FUNCTION_BLOCK "FB_SatelliteUnit"   // FB4, SCL
{ S7_Optimized_Access := 'TRUE' }
VERSION : 0.1
// Generated frame v0.12; change the declaration, then regenerate.
// stored: AutoNumber true, IsIECCheckEnabled false, IsRetainMemResEnabled false, MemoryReserve 100, SetENOAutomatically false, UDAEnableTagReadback false
   VAR_INPUT
      Execute { ExternalWritable := 'False'} : Bool;
      Abort { ExternalWritable := 'False'} : Bool;
      Command { ExternalWritable := 'False'} : DInt;
      ParCmd { ExternalWritable := 'False'} : "ST_DeclarationParCmd";
      ParentIndex { ExternalAccessible := 'False'; ExternalVisible := 'False'; ExternalWritable := 'False'} : DInt;
      Startup { ExternalAccessible := 'False'; ExternalVisible := 'False'; ExternalWritable := 'False'} : Bool;
   END_VAR
   VAR_OUTPUT
      Busy { ExternalWritable := 'False'} : Bool;
      Done { ExternalWritable := 'False'} : Bool;
      Error { ExternalWritable := 'False'} : Bool;
      Aborted { ExternalWritable := 'False'} : Bool;
      Held { ExternalWritable := 'False'} : Bool;
      ErrorID { ExternalWritable := 'False'} : DWord;
      Timing { ExternalWritable := 'False'} : "ST_ModuleTiming";
      OutCmd { ExternalWritable := 'False'} : "ST_DeclarationOutCmd";
      OutImm { ExternalWritable := 'False'} : "ST_UnitProbeImm";
   END_VAR
   VAR_IN_OUT
      Hal : "ST_SatelliteUnitHal";
   END_VAR
   VAR
      Status { ExternalWritable := 'False'; S7_SetPoint := 'True'} : "ST_ModuleStatus";
      Core { ExternalAccessible := 'False'; ExternalVisible := 'False'; ExternalWritable := 'False'; S7_SetPoint := 'True'} : "FRK_Core";
      ParCfg { ExternalWritable := 'False'; S7_SetPoint := 'True'} : "ST_DeclarationParCfg";
      LatchedParCmd { ExternalAccessible := 'False'; ExternalVisible := 'False'; ExternalWritable := 'False'; S7_SetPoint := 'True'} : "ST_DeclarationParCmd";
      StateFlags { ExternalWritable := 'False'; S7_SetPoint := 'True'} : Array[1..12] of "ST_StateFlag";
      StateFlagCount { ExternalWritable := 'False'} : Int;
      StateTouched { ExternalAccessible := 'False'; ExternalVisible := 'False'; ExternalWritable := 'False'} : Array[1..12] of Bool;
      Device { ExternalAccessible := 'False'; ExternalVisible := 'False'; ExternalWritable := 'False'; S7_SetPoint := 'True'} : "ST_UnitProbeDevice";
      StationCfg { ExternalWritable := 'False'; S7_SetPoint := 'True'} : "ST_UnitProbeStationCfg";
      ConfigStageParCfg { ExternalAccessible := 'False'; ExternalVisible := 'False'; ExternalWritable := 'False'; S7_SetPoint := 'True'} : "ST_DeclarationParCfg";
      ConfigDefaultParCfg { ExternalAccessible := 'False'; ExternalVisible := 'False'; ExternalWritable := 'False'; S7_SetPoint := 'True'} : "ST_DeclarationParCfg";
      ConfigStageStationCfg { ExternalAccessible := 'False'; ExternalVisible := 'False'; ExternalWritable := 'False'; S7_SetPoint := 'True'} : "ST_UnitProbeStationCfg";
      ConfigDefaultStationCfg { ExternalAccessible := 'False'; ExternalVisible := 'False'; ExternalWritable := 'False'; S7_SetPoint := 'True'} : "ST_UnitProbeStationCfg";
      ConfigStaged { ExternalAccessible := 'False'; ExternalVisible := 'False'; ExternalWritable := 'False'} : Bool;
      Unit { ExternalAccessible := 'False'; ExternalVisible := 'False'; ExternalWritable := 'False'; S7_SetPoint := 'True'} : "FRK_Unit";
      HmiRequest { S7_SetPoint := 'True'} : "ST_HmiRequest";
      ModePolicy { ExternalAccessible := 'False'; ExternalVisible := 'False'; ExternalWritable := 'False'; S7_SetPoint := 'True'} : Array[0..6] of "ST_ModePolicy";
      Access { ExternalWritable := 'False'; S7_SetPoint := 'True'} : "FRK_Access";
      HmiResponse { ExternalWritable := 'False'; S7_SetPoint := 'True'} : "ST_HmiResponse";
      ConfigRev { ExternalWritable := 'False'} : UDInt;
      ConfigCursor { ExternalAccessible := 'False'; ExternalVisible := 'False'; ExternalWritable := 'False'; S7_SetPoint := 'True'} : "FRK_ConfigCursor";
      Part { ExternalWritable := 'False'; S7_SetPoint := 'True'} : "ST_PartContext";
      Decision { ExternalWritable := 'False'; S7_SetPoint := 'True'} : "ST_DecisionRequest";
      DecisionAnswer { ExternalWritable := 'False'} : Int;
      History { ExternalWritable := 'False'; S7_SetPoint := 'True'} : Array[1..16] of "ST_Diagnostic";
      HistoryHead { ExternalWritable := 'False'} : Int;
      AlarmLog { ExternalWritable := 'False'; S7_SetPoint := 'True'} : "FRK_AlarmLog";
      ModeActivePublished { ExternalWritable := 'False'} : DInt;
      RunningPublished { ExternalWritable := 'False'} : Bool;
      StopPendingPublished { ExternalWritable := 'False'} : Bool;
      SupportedModesPublished { ExternalWritable := 'False'} : Array[0..6] of Bool;
      GoodCount { ExternalWritable := 'False'} : UDInt;
      NokCount { ExternalWritable := 'False'} : UDInt;
      ReworkCount { ExternalWritable := 'False'} : UDInt;
      NokReason { ExternalWritable := 'False'} : DInt;
      Cell { ExternalWritable := 'False'; S7_SetPoint := 'True'} : "FB_DeclarationCell";
      Inner { ExternalWritable := 'False'; S7_SetPoint := 'True'} : "FB_InnerUnit";
   END_VAR
   VAR_TEMP
      InstancePath : WString[254];
      RouteMatched : Bool;
      ManualMatched : Bool;
   END_VAR
   VAR CONSTANT
      EXEC_READY : DInt := 0;
      MODULE_TIER : DInt := 1;
   END_VAR
BEGIN

   // ---- GENERATED: setup
   IF #Startup OR NOT #Core.Named THEN
       #InstancePath := GetInstancePath(size := 0);
       "FRK_SetIdentity"(Core := #Core,
                         Status := #Status,
                         InstancePath := #InstancePath,
                         ModuleType := 1,
                         TypeId := 4,
                         Capabilities := DWORD#16#00000000,
                         ParentIndex := #ParentIndex,
                         TypeKey := 'Fraktal.Test.Satellite');
   END_IF;
   IF #Startup THEN "FRK_CfgRestore_SatelliteUnit"(Core := #Core,
                                                       Status := #Status,
                                                       ParCfg := #ParCfg,
                                                       StationCfg := #StationCfg,
                                                       ConfigStageParCfg := #ConfigStageParCfg,
                                                       ConfigDefaultParCfg := #ConfigDefaultParCfg,
                                                       ConfigStageStationCfg := #ConfigStageStationCfg,
                                                       ConfigDefaultStationCfg := #ConfigDefaultStationCfg);
   END_IF;
   "FRK_StateSweep"(Flags := #StateFlags,
                    Count := #StateFlagCount,
                    Touched := #StateTouched,
                    Startup := #Startup);
   IF #Startup OR #ConfigRev = 0 THEN
       #ConfigRev := "FRK_ConfigRevision"(Previous := #ConfigRev);
   END_IF;
   #SupportedModesPublished[0] := TRUE;
   #SupportedModesPublished[1] := TRUE;
   #SupportedModesPublished[2] := TRUE;
   #SupportedModesPublished[3] := FALSE;
   #SupportedModesPublished[4] := FALSE;
   #SupportedModesPublished[5] := FALSE;
   #SupportedModesPublished[6] := FALSE;
   "FRK_UnitPrepare"(Core := #Core,
                     Unit := #Unit,
                     Policy := #ModePolicy,
                     Request := #HmiRequest,
                     Response := #HmiResponse,
                     Startup := #Startup,
                     InitialMode := 1);
   "FRK_AlarmBegin"(AlarmLog := #AlarmLog,
                    Startup := #Startup);
   "FRK_AlarmHistoryBoot"(AlarmLog := #AlarmLog,
                          Startup := #Startup,
                          Scope := #Status.Name);
   "FRK_AccessPolicyBoot"(Access := #Access,
                          Startup := #Startup,
                          Root := #Core.ParentIndex = 0,
                          Scope := #Status.Name);
   "FRK_AccessCyclic"(Access := #Access,
                      Startup := #Startup,
                      SourcePath := STRING_TO_WSTRING(#Status.Name),
                      AlarmLog := #AlarmLog,
                      Revision := #ConfigRev);
   "FRK_UnitMailbox"(Core := #Core,
                     Unit := #Unit,
                     Status := #Status,
                     Policy := #ModePolicy,
                     Access := #Access,
                     Request := #HmiRequest,
                     Response := #HmiResponse,
                     Supported := #SupportedModesPublished);
   #Unit.ConfigBlocked := #Access.PolicyLost;
   // ---- GENERATED: begin
   "FRK_Begin"(Core := #Core,
               Status := #Status,
               Execute := #Unit.RunReq,
               Abort := (#Abort OR #Unit.AbortReq),
               Command := 1);
   IF #Core.EvCommandStart THEN
       #LatchedParCmd := #ParCmd;
       CASE #Core.Command OF
           1:
               "FRK_UnitRunStart"(Core := #Core,
                                  Status := #Status,
                                  Timeout := #ParCfg.Timeout,
                                  Label := 'Run');
           ELSE
               "FRK_Start"(Core := #Core,
                           Status := #Status,
                           Supported := FALSE,
                           Timeout := T#0ms,
                           Label := '');
       END_CASE;
   END_IF;
   IF #Core.EvCommandStart THEN
       // ---- AUTHORED: CommandStart
       #Device.Received := "FRK_PartReceived"(Core := #Core, Unit := #Unit, Status := #Status, Part := #Part, AlarmLog := #AlarmLog);
       IF #Device.Received THEN
           "FRK_PartStarted"(Unit := #Unit,
                             Status := #Status,
                             Part := #Part,
                             AlarmLog := #AlarmLog);
       END_IF;
       // ---- GENERATED: reaction end
   END_IF;
   // ---- AUTHORED: cyclic management
   IF #Hal.Cell.Clamp.BackgroundFault THEN
       "FRK_Fault"(Core := #Core,
                   Status := #Status,
                   ReasonCode := 2901,
                   Description := WSTRING#'test.unit.condition');
   END_IF;
   // ---- GENERATED: end management
   "FRK_Release_SatelliteUnit"(Unit := #Unit,
                               Hal := #Hal);
   IF #Core.RegIndex > 0 THEN
       "FRK_Registry".Rows[#Core.RegIndex].AlarmBlocking := #AlarmLog.Blocking;
   END_IF;
   #Unit.AlarmBlocking := "FRK_AlarmTreeBlocking"(Owner := #Core.RegIndex);
   "FRK_UnitConsume"(Core := #Core,
                     Unit := #Unit,
                     Status := #Status,
                     Policy := #ModePolicy,
                     Access := #Access,
                     Response := #HmiResponse,
                     Supported := #SupportedModesPublished);
   "FRK_UnitMode"(Core := #Core,
                  Unit := #Unit);
   IF #Core.EvModeExit THEN
       // ---- AUTHORED: ModeExit
       #Device.ExitCalls := #Device.ExitCalls + 1;
       IF #Hal.Cell.Clamp.ExitHold THEN
           #Core.HookResult := 1;
       ELSE
           #Core.HookResult := 0;
       END_IF;
       // ---- GENERATED: reaction end
   END_IF;
   "FRK_UnitModeResolve"(Core := #Core,
                         Unit := #Unit,
                         Status := #Status,
                         Policy := #ModePolicy,
                         Timeout := #ParCfg.Timeout);
   IF #Core.EvModeChanged THEN
       // ---- AUTHORED: ModeChanged
       #Device.Changes := #Device.Changes + 1;
       // ---- GENERATED: reaction end
   END_IF;
   "FRK_DecisionCyclic"(Owner := #Core.RegIndex,
                        Busy := #Core.Exec = 1,
                        Reset := #Startup OR #Unit.EvReset OR #Core.EvModeChanged,
                        AlarmLog := #AlarmLog);
   "FRK_UnitFollow"(Core := #Core,
                    Unit := #Unit,
                    Status := #Status,
                    Policy := #ModePolicy,
                    Access := #Access,
                    Supported := #SupportedModesPublished);
   IF #Unit.RequestPending AND (#Unit.Request.Kind = 11 OR #Unit.Request.Kind = 16) THEN
       #ManualMatched := FALSE;
       #RouteMatched := "FRK_Route_DeclarationCell"(Module := #Cell, Hal := #Hal.Cell, Request := #Unit.Request, Report := #HmiResponse.Report);
       #ManualMatched := #ManualMatched OR #RouteMatched;
       #RouteMatched := "FRK_Route_InnerUnit"(Module := #Inner, Hal := #Hal.Inner, Request := #Unit.Request, Report := #HmiResponse.Report);
       #ManualMatched := #ManualMatched OR #RouteMatched;
       IF NOT #ManualMatched THEN
           "FRK_ReleaseReason"(Report := #HmiResponse.Report,
                               Description := WSTRING#'std.error.unsupportedHmiRequest',
                               Reason := 2008,
                               Path := #Unit.Request.TargetPath,
                               Kind := 4);
       END_IF;
       #HmiResponse.Accepted := #Unit.Request.Kind = 16 OR #HmiResponse.Report.Released;
       IF #Unit.Request.Kind = 11 THEN
           IF #HmiResponse.Accepted THEN
               #HmiResponse.Diagnostic := WSTRING#'std.audit.manualCommandAccepted';
           ELSE
               #HmiResponse.Diagnostic := WSTRING#'std.audit.manualCommandRejected';
           END_IF;
       END_IF;
   END_IF;
   IF #Unit.EvReset THEN
       "FRK_AlarmOperatorReset"(AlarmLog := #AlarmLog);
   END_IF;
   IF #Unit.EvReset THEN
       // ---- AUTHORED: OperatorReset
       #Device.Resets := #Device.Resets + 1;
       // ---- GENERATED: reset reaction end
   END_IF;
   IF #Core.ReleasePending OR #Unit.ReleaseChildren THEN
       "FRK_ReleaseCommand"(Core := #Cell.Core,
                            Execute := #Cell.Execute);
       "FRK_ReleaseCommand"(Core := #Inner.Core,
                            Execute := #Inner.Execute);
   END_IF;
   // ---- GENERATED: child call
   #Cell(ParentIndex := #Core.RegIndex,
         Startup := #Startup,
         Hal := #Hal.Cell);
   "FRK_ManualFinish"(Core := #Cell.Core,
                      Execute := #Cell.Execute,
                      ManualOwned := #Cell.ManualOwned);
   "FRK_UnitCascade"(ParentUnit := #Unit,
                     Core := #Inner.Core,
                     Unit := #Inner.Unit,
                     Status := #Inner.Status,
                     Policy := #Inner.ModePolicy,
                     Access := #Inner.Access,
                     Supported := #Inner.SupportedModesPublished,
                     AlarmLog := #AlarmLog);
   // ---- GENERATED: child call
   #Inner(ParentIndex := #Core.RegIndex,
          Startup := #Startup,
          Hal := #Hal.Inner);
   #Unit.CascadePending := FALSE;
   IF #Unit.RequestPending AND #Unit.Request.Kind = 23 THEN
       #HmiResponse.Accepted := FALSE;
       #HmiResponse.Report.Count := 0;
       #HmiResponse.Report.Released := TRUE;
       #HmiResponse.Diagnostic := WSTRING#'';
       "FRK_ConfigBegin"(Cursor := #ConfigCursor,
                         Page := #HmiResponse.ConfigPage,
                         PageIndex := #Unit.Request.IntValue,
                         Revision := #ConfigRev);
       IF #Unit.Request.DurationMs <> 0 THEN
           #HmiResponse.Diagnostic := WSTRING#'std.error.modelNotAvailable';
       ELSIF #Unit.Request.IntValue < 0 OR #Unit.Request.IntValue > 32767 THEN
           #HmiResponse.Diagnostic := WSTRING#'std.error.hmiRequestRejected';
       ELSE
           "FRK_ConfigUnit"(Scope := #Status.Name,
                            Policy := #ModePolicy,
                            ModelCount := 0,
                            ReadLevel := #Access.Policy.Required[0],
                            Readable := #Access.CurrentLevel >= #Access.Policy.Required[0],
                            Cursor := #ConfigCursor,
                            Page := #HmiResponse.ConfigPage);
           "FRK_Config_DeclarationCell"(Module := #Cell,
                                        Access := #Access,
                                        RootIndex := "FRK_ConfigRoot"(RegIndex := #Core.RegIndex),
                                        ModelIndex := 0,
                                        Cursor := #ConfigCursor,
                                        Page := #HmiResponse.ConfigPage);
           "FRK_Config_InnerUnit"(Module := #Inner,
                                  Access := #Access,
                                  RootIndex := "FRK_ConfigRoot"(RegIndex := #Core.RegIndex),
                                  ModelIndex := 0,
                                  Cursor := #ConfigCursor,
                                  Page := #HmiResponse.ConfigPage);
           "FRK_ConfigFinish"(Cursor := #ConfigCursor,
                              Page := #HmiResponse.ConfigPage);
           #HmiResponse.Accepted := TRUE;
       END_IF;
   END_IF;
   "FRK_RouteAbort"(Core := #Core,
                    Abort := (#Abort OR #Unit.AbortReq));
   IF #Core.EvAbort THEN
       "FRK_PartAborted"(Core := #Core,
                         Unit := #Unit,
                         Status := #Status,
                         Part := #Part,
                         AlarmLog := #AlarmLog);
   END_IF;
   IF #Core.Dispatch AND #Core.RegIndex > 0 AND NOT "FRK_Registry".Fault THEN
       // ---- AUTHORED: dispatch
       IF #Hal.Cell.Clamp.Finish THEN
           #Device.Processed := FALSE;
           IF #Unit.CarrierIndex = 0 THEN
               #Device.Processed := TRUE;
           ELSE
               #Device.Processed := "FRK_PartProcessed"(Core := #Core, Unit := #Unit, Status := #Status, Part := #Part, AlarmLog := #AlarmLog, Verdict := #Hal.Cell.Clamp.Verdict, Reason := #Hal.Cell.Clamp.Diag.ReasonCode);
           END_IF;
           IF #Device.Processed THEN
               #Device.Cycles := #Device.Cycles + 1;
               IF #Unit.StopReq THEN
                   "FRK_Complete"(Core := #Core,
                                  Status := #Status);
               ELSE
                   #Device.Received := "FRK_PartReceived"(Core := #Core, Unit := #Unit, Status := #Status, Part := #Part, AlarmLog := #AlarmLog);
                   IF #Device.Received THEN
                       "FRK_PartStarted"(Unit := #Unit,
                                         Status := #Status,
                                         Part := #Part,
                                         AlarmLog := #AlarmLog);
                   END_IF;
               END_IF;
           END_IF;
       END_IF;
       // ---- GENERATED: end dispatch
   END_IF;
   "FRK_End"(Core := #Core,
             Status := #Status,
             Busy => #Busy,
             Done => #Done,
             Error => #Error,
             Aborted => #Aborted,
             Held => #Held,
             ErrorID => #ErrorID,
             Timing => #Timing);
   "FRK_DecisionCyclic"(Owner := #Core.RegIndex,
                        Busy := #Core.Exec = 1,
                        Reset := #Startup OR #Unit.EvReset OR #Core.EvModeChanged,
                        AlarmLog := #AlarmLog);
   "FRK_DecisionPublish"(Owner := #Core.RegIndex,
                         Decision := #Decision,
                         DecisionAnswer := #DecisionAnswer);
   IF NOT #Unit.EvReset THEN
       "FRK_AlarmCapture"(AlarmLog := #AlarmLog,
                          Core := #Core,
                          Status := #Status);
       "FRK_Capture_DeclarationCell"(Module := #Cell,
                                     AlarmLog := #AlarmLog);
       "FRK_AlarmEnd"(AlarmLog := #AlarmLog);
   END_IF;
   IF #Core.RegIndex > 0 THEN
       "FRK_Registry".Rows[#Core.RegIndex].AlarmBlocking := #AlarmLog.Blocking;
   END_IF;
   #Unit.AlarmBlocking := "FRK_AlarmTreeBlocking"(Owner := #Core.RegIndex);
   "FRK_AccessPersist"(Access := #Access,
                       Unit := #Unit,
                       Response := #HmiResponse,
                       SourcePath := STRING_TO_WSTRING(#Status.Name),
                       AlarmLog := #AlarmLog);
   "FRK_AccessFinish"(Access := #Access,
                      Unit := #Unit,
                      Response := #HmiResponse,
                      SourcePath := STRING_TO_WSTRING(#Status.Name),
                      AlarmLog := #AlarmLog,
                      Revision := #ConfigRev);
   "FRK_UnitFinish"(Core := #Core,
                    Unit := #Unit,
                    Response := #HmiResponse,
                    Status := #Status,
                    Part := #Part,
                    AlarmLog := #AlarmLog,
                    History := #History,
                    Head := #HistoryHead);
   #ModeActivePublished := #Unit.Mode;
   #RunningPublished := #Core.Exec = 1;
   #StopPendingPublished := #Unit.StopReq AND #Core.Exec = 1;
   #GoodCount := #Unit.Good;
   #NokCount := #Unit.Nok;
   #ReworkCount := #Unit.Rework;
   #NokReason := #Unit.NokReason;
   // ---- AUTHORED: unconditional cyclic/derived data
   #OutImm.Cycles := #Device.Cycles;
   #OutImm.ExitCalls := #Device.ExitCalls;
   #OutImm.Changes := #Device.Changes;
   #OutImm.Resets := #Device.Resets;
   #OutImm.AtHome := "FRK_State"(Idx := 1, Key := 'project.state.atHome', Ok := #Hal.Cell.Clamp.Sample = 0, Flags := #StateFlags, Count := #StateFlagCount, Touched := #StateTouched);
   // ---- GENERATED: frame end
END_FUNCTION_BLOCK

FUNCTION_BLOCK "FB_InnerUnit"   // FB3, SCL
{ S7_Optimized_Access := 'TRUE' }
VERSION : 0.1
// Generated frame v0.12; change the declaration, then regenerate.
// stored: AutoNumber true, IsIECCheckEnabled false, IsRetainMemResEnabled false, MemoryReserve 100, SetENOAutomatically false, UDAEnableTagReadback false
   VAR_INPUT
      Execute { ExternalWritable := 'False'} : Bool;
      Abort { ExternalWritable := 'False'} : Bool;
      Command { ExternalWritable := 'False'} : DInt;
      ParCmd { ExternalWritable := 'False'} : "ST_DeclarationParCmd";
      ParentIndex { ExternalAccessible := 'False'; ExternalVisible := 'False'; ExternalWritable := 'False'} : DInt;
      Startup { ExternalAccessible := 'False'; ExternalVisible := 'False'; ExternalWritable := 'False'} : Bool;
   END_VAR
   VAR_OUTPUT
      Busy { ExternalWritable := 'False'} : Bool;
      Done { ExternalWritable := 'False'} : Bool;
      Error { ExternalWritable := 'False'} : Bool;
      Aborted { ExternalWritable := 'False'} : Bool;
      Held { ExternalWritable := 'False'} : Bool;
      ErrorID { ExternalWritable := 'False'} : DWord;
      Timing { ExternalWritable := 'False'} : "ST_ModuleTiming";
      OutCmd { ExternalWritable := 'False'} : "ST_DeclarationOutCmd";
      OutImm { ExternalWritable := 'False'} : "ST_UnitProbeImm";
   END_VAR
   VAR_IN_OUT
      Hal : "ST_InnerUnitHal";
   END_VAR
   VAR
      Status { ExternalWritable := 'False'; S7_SetPoint := 'True'} : "ST_ModuleStatus";
      Core { ExternalAccessible := 'False'; ExternalVisible := 'False'; ExternalWritable := 'False'; S7_SetPoint := 'True'} : "FRK_Core";
      ParCfg { ExternalWritable := 'False'; S7_SetPoint := 'True'} : "ST_DeclarationParCfg";
      LatchedParCmd { ExternalAccessible := 'False'; ExternalVisible := 'False'; ExternalWritable := 'False'; S7_SetPoint := 'True'} : "ST_DeclarationParCmd";
      StateFlags { ExternalWritable := 'False'; S7_SetPoint := 'True'} : Array[1..12] of "ST_StateFlag";
      StateFlagCount { ExternalWritable := 'False'} : Int;
      StateTouched { ExternalAccessible := 'False'; ExternalVisible := 'False'; ExternalWritable := 'False'} : Array[1..12] of Bool;
      Device { ExternalAccessible := 'False'; ExternalVisible := 'False'; ExternalWritable := 'False'; S7_SetPoint := 'True'} : "ST_UnitProbeDevice";
      StationCfg { ExternalWritable := 'False'; S7_SetPoint := 'True'} : "ST_UnitProbeStationCfg";
      ConfigStageParCfg { ExternalAccessible := 'False'; ExternalVisible := 'False'; ExternalWritable := 'False'; S7_SetPoint := 'True'} : "ST_DeclarationParCfg";
      ConfigDefaultParCfg { ExternalAccessible := 'False'; ExternalVisible := 'False'; ExternalWritable := 'False'; S7_SetPoint := 'True'} : "ST_DeclarationParCfg";
      ConfigStageStationCfg { ExternalAccessible := 'False'; ExternalVisible := 'False'; ExternalWritable := 'False'; S7_SetPoint := 'True'} : "ST_UnitProbeStationCfg";
      ConfigDefaultStationCfg { ExternalAccessible := 'False'; ExternalVisible := 'False'; ExternalWritable := 'False'; S7_SetPoint := 'True'} : "ST_UnitProbeStationCfg";
      ConfigStaged { ExternalAccessible := 'False'; ExternalVisible := 'False'; ExternalWritable := 'False'} : Bool;
      Unit { ExternalAccessible := 'False'; ExternalVisible := 'False'; ExternalWritable := 'False'; S7_SetPoint := 'True'} : "FRK_Unit";
      HmiRequest { S7_SetPoint := 'True'} : "ST_HmiRequest";
      ModePolicy { ExternalAccessible := 'False'; ExternalVisible := 'False'; ExternalWritable := 'False'; S7_SetPoint := 'True'} : Array[0..6] of "ST_ModePolicy";
      Access { ExternalWritable := 'False'; S7_SetPoint := 'True'} : "FRK_Access";
      HmiResponse { ExternalWritable := 'False'; S7_SetPoint := 'True'} : "ST_HmiResponse";
      ConfigRev { ExternalWritable := 'False'} : UDInt;
      ConfigCursor { ExternalAccessible := 'False'; ExternalVisible := 'False'; ExternalWritable := 'False'; S7_SetPoint := 'True'} : "FRK_ConfigCursor";
      Part { ExternalWritable := 'False'; S7_SetPoint := 'True'} : "ST_PartContext";
      Decision { ExternalWritable := 'False'; S7_SetPoint := 'True'} : "ST_DecisionRequest";
      DecisionAnswer { ExternalWritable := 'False'} : Int;
      History { ExternalWritable := 'False'; S7_SetPoint := 'True'} : Array[1..16] of "ST_Diagnostic";
      HistoryHead { ExternalWritable := 'False'} : Int;
      AlarmLog { ExternalWritable := 'False'; S7_SetPoint := 'True'} : "FRK_AlarmLog";
      ModeActivePublished { ExternalWritable := 'False'} : DInt;
      RunningPublished { ExternalWritable := 'False'} : Bool;
      StopPendingPublished { ExternalWritable := 'False'} : Bool;
      SupportedModesPublished { ExternalWritable := 'False'} : Array[0..6] of Bool;
      GoodCount { ExternalWritable := 'False'} : UDInt;
      NokCount { ExternalWritable := 'False'} : UDInt;
      ReworkCount { ExternalWritable := 'False'} : UDInt;
      NokReason { ExternalWritable := 'False'} : DInt;
      Cell { ExternalWritable := 'False'; S7_SetPoint := 'True'} : "FB_DeclarationCell";
   END_VAR
   VAR_TEMP
      InstancePath : WString[254];
      RouteMatched : Bool;
      ManualMatched : Bool;
   END_VAR
   VAR CONSTANT
      EXEC_READY : DInt := 0;
      MODULE_TIER : DInt := 1;
   END_VAR
BEGIN

   // ---- GENERATED: setup
   IF #Startup OR NOT #Core.Named THEN
       #InstancePath := GetInstancePath(size := 0);
       "FRK_SetIdentity"(Core := #Core,
                         Status := #Status,
                         InstancePath := #InstancePath,
                         ModuleType := 1,
                         TypeId := 5,
                         Capabilities := DWORD#16#00000000,
                         ParentIndex := #ParentIndex,
                         TypeKey := 'Fraktal.Test.Inner');
   END_IF;
   IF #Startup THEN "FRK_CfgRestore_InnerUnit"(Core := #Core,
                                                   Status := #Status,
                                                   ParCfg := #ParCfg,
                                                   StationCfg := #StationCfg,
                                                   ConfigStageParCfg := #ConfigStageParCfg,
                                                   ConfigDefaultParCfg := #ConfigDefaultParCfg,
                                                   ConfigStageStationCfg := #ConfigStageStationCfg,
                                                   ConfigDefaultStationCfg := #ConfigDefaultStationCfg);
   END_IF;
   "FRK_StateSweep"(Flags := #StateFlags,
                    Count := #StateFlagCount,
                    Touched := #StateTouched,
                    Startup := #Startup);
   IF #Startup OR #ConfigRev = 0 THEN
       #ConfigRev := "FRK_ConfigRevision"(Previous := #ConfigRev);
   END_IF;
   #SupportedModesPublished[0] := TRUE;
   #SupportedModesPublished[1] := TRUE;
   #SupportedModesPublished[2] := TRUE;
   #SupportedModesPublished[3] := FALSE;
   #SupportedModesPublished[4] := FALSE;
   #SupportedModesPublished[5] := FALSE;
   #SupportedModesPublished[6] := FALSE;
   "FRK_UnitPrepare"(Core := #Core,
                     Unit := #Unit,
                     Policy := #ModePolicy,
                     Request := #HmiRequest,
                     Response := #HmiResponse,
                     Startup := #Startup,
                     InitialMode := 1);
   "FRK_AlarmBegin"(AlarmLog := #AlarmLog,
                    Startup := #Startup);
   "FRK_AlarmHistoryBoot"(AlarmLog := #AlarmLog,
                          Startup := #Startup,
                          Scope := #Status.Name);
   "FRK_AccessPolicyBoot"(Access := #Access,
                          Startup := #Startup,
                          Root := #Core.ParentIndex = 0,
                          Scope := #Status.Name);
   "FRK_AccessCyclic"(Access := #Access,
                      Startup := #Startup,
                      SourcePath := STRING_TO_WSTRING(#Status.Name),
                      AlarmLog := #AlarmLog,
                      Revision := #ConfigRev);
   "FRK_UnitMailbox"(Core := #Core,
                     Unit := #Unit,
                     Status := #Status,
                     Policy := #ModePolicy,
                     Access := #Access,
                     Request := #HmiRequest,
                     Response := #HmiResponse,
                     Supported := #SupportedModesPublished);
   #Unit.ConfigBlocked := #Access.PolicyLost;
   // ---- GENERATED: begin
   "FRK_Begin"(Core := #Core,
               Status := #Status,
               Execute := #Unit.RunReq,
               Abort := (#Abort OR #Unit.AbortReq),
               Command := 1);
   IF #Core.EvCommandStart THEN
       #LatchedParCmd := #ParCmd;
       CASE #Core.Command OF
           1:
               "FRK_UnitRunStart"(Core := #Core,
                                  Status := #Status,
                                  Timeout := #ParCfg.Timeout,
                                  Label := 'Run');
           ELSE
               "FRK_Start"(Core := #Core,
                           Status := #Status,
                           Supported := FALSE,
                           Timeout := T#0ms,
                           Label := '');
       END_CASE;
   END_IF;
   IF #Core.EvCommandStart THEN
       // ---- AUTHORED: CommandStart
       #Device.Received := "FRK_PartReceived"(Core := #Core, Unit := #Unit, Status := #Status, Part := #Part, AlarmLog := #AlarmLog);
       IF #Device.Received THEN
           "FRK_PartStarted"(Unit := #Unit,
                             Status := #Status,
                             Part := #Part,
                             AlarmLog := #AlarmLog);
       END_IF;
       // ---- GENERATED: reaction end
   END_IF;
   // ---- AUTHORED: cyclic management
   IF #Hal.Cell.Clamp.BackgroundFault THEN
       "FRK_Fault"(Core := #Core,
                   Status := #Status,
                   ReasonCode := 2901,
                   Description := WSTRING#'test.unit.condition');
   END_IF;
   // ---- GENERATED: end management
   "FRK_Release_InnerUnit"(Unit := #Unit,
                           Hal := #Hal);
   IF #Core.RegIndex > 0 THEN
       "FRK_Registry".Rows[#Core.RegIndex].AlarmBlocking := #AlarmLog.Blocking;
   END_IF;
   #Unit.AlarmBlocking := "FRK_AlarmTreeBlocking"(Owner := #Core.RegIndex);
   "FRK_UnitConsume"(Core := #Core,
                     Unit := #Unit,
                     Status := #Status,
                     Policy := #ModePolicy,
                     Access := #Access,
                     Response := #HmiResponse,
                     Supported := #SupportedModesPublished);
   "FRK_UnitMode"(Core := #Core,
                  Unit := #Unit);
   IF #Core.EvModeExit THEN
       // ---- AUTHORED: ModeExit
       #Device.ExitCalls := #Device.ExitCalls + 1;
       IF #Hal.Cell.Clamp.ExitHold THEN
           #Core.HookResult := 1;
       ELSE
           #Core.HookResult := 0;
       END_IF;
       // ---- GENERATED: reaction end
   END_IF;
   "FRK_UnitModeResolve"(Core := #Core,
                         Unit := #Unit,
                         Status := #Status,
                         Policy := #ModePolicy,
                         Timeout := #ParCfg.Timeout);
   IF #Core.EvModeChanged THEN
       // ---- AUTHORED: ModeChanged
       #Device.Changes := #Device.Changes + 1;
       // ---- GENERATED: reaction end
   END_IF;
   "FRK_DecisionCyclic"(Owner := #Core.RegIndex,
                        Busy := #Core.Exec = 1,
                        Reset := #Startup OR #Unit.EvReset OR #Core.EvModeChanged,
                        AlarmLog := #AlarmLog);
   "FRK_UnitFollow"(Core := #Core,
                    Unit := #Unit,
                    Status := #Status,
                    Policy := #ModePolicy,
                    Access := #Access,
                    Supported := #SupportedModesPublished);
   IF #Unit.RequestPending AND (#Unit.Request.Kind = 11 OR #Unit.Request.Kind = 16) THEN
       #ManualMatched := FALSE;
       #RouteMatched := "FRK_Route_DeclarationCell"(Module := #Cell, Hal := #Hal.Cell, Request := #Unit.Request, Report := #HmiResponse.Report);
       #ManualMatched := #ManualMatched OR #RouteMatched;
       IF NOT #ManualMatched THEN
           "FRK_ReleaseReason"(Report := #HmiResponse.Report,
                               Description := WSTRING#'std.error.unsupportedHmiRequest',
                               Reason := 2008,
                               Path := #Unit.Request.TargetPath,
                               Kind := 4);
       END_IF;
       #HmiResponse.Accepted := #Unit.Request.Kind = 16 OR #HmiResponse.Report.Released;
       IF #Unit.Request.Kind = 11 THEN
           IF #HmiResponse.Accepted THEN
               #HmiResponse.Diagnostic := WSTRING#'std.audit.manualCommandAccepted';
           ELSE
               #HmiResponse.Diagnostic := WSTRING#'std.audit.manualCommandRejected';
           END_IF;
       END_IF;
   END_IF;
   IF #Unit.EvReset THEN
       "FRK_AlarmOperatorReset"(AlarmLog := #AlarmLog);
   END_IF;
   IF #Unit.EvReset THEN
       // ---- AUTHORED: OperatorReset
       #Device.Resets := #Device.Resets + 1;
       // ---- GENERATED: reset reaction end
   END_IF;
   IF #Core.ReleasePending OR #Unit.ReleaseChildren THEN
       "FRK_ReleaseCommand"(Core := #Cell.Core,
                            Execute := #Cell.Execute);
   END_IF;
   // ---- GENERATED: child call
   #Cell(ParentIndex := #Core.RegIndex,
         Startup := #Startup,
         Hal := #Hal.Cell);
   "FRK_ManualFinish"(Core := #Cell.Core,
                      Execute := #Cell.Execute,
                      ManualOwned := #Cell.ManualOwned);
   #Unit.CascadePending := FALSE;
   IF #Unit.RequestPending AND #Unit.Request.Kind = 23 THEN
       #HmiResponse.Accepted := FALSE;
       #HmiResponse.Report.Count := 0;
       #HmiResponse.Report.Released := TRUE;
       #HmiResponse.Diagnostic := WSTRING#'';
       "FRK_ConfigBegin"(Cursor := #ConfigCursor,
                         Page := #HmiResponse.ConfigPage,
                         PageIndex := #Unit.Request.IntValue,
                         Revision := #ConfigRev);
       IF #Unit.Request.DurationMs <> 0 THEN
           #HmiResponse.Diagnostic := WSTRING#'std.error.modelNotAvailable';
       ELSIF #Unit.Request.IntValue < 0 OR #Unit.Request.IntValue > 32767 THEN
           #HmiResponse.Diagnostic := WSTRING#'std.error.hmiRequestRejected';
       ELSE
           "FRK_ConfigUnit"(Scope := #Status.Name,
                            Policy := #ModePolicy,
                            ModelCount := 0,
                            ReadLevel := #Access.Policy.Required[0],
                            Readable := #Access.CurrentLevel >= #Access.Policy.Required[0],
                            Cursor := #ConfigCursor,
                            Page := #HmiResponse.ConfigPage);
           "FRK_Config_DeclarationCell"(Module := #Cell,
                                        Access := #Access,
                                        RootIndex := "FRK_ConfigRoot"(RegIndex := #Core.RegIndex),
                                        ModelIndex := 0,
                                        Cursor := #ConfigCursor,
                                        Page := #HmiResponse.ConfigPage);
           "FRK_ConfigFinish"(Cursor := #ConfigCursor,
                              Page := #HmiResponse.ConfigPage);
           #HmiResponse.Accepted := TRUE;
       END_IF;
   END_IF;
   "FRK_RouteAbort"(Core := #Core,
                    Abort := (#Abort OR #Unit.AbortReq));
   IF #Core.EvAbort THEN
       "FRK_PartAborted"(Core := #Core,
                         Unit := #Unit,
                         Status := #Status,
                         Part := #Part,
                         AlarmLog := #AlarmLog);
   END_IF;
   IF #Core.Dispatch AND #Core.RegIndex > 0 AND NOT "FRK_Registry".Fault THEN
       // ---- AUTHORED: dispatch
       IF #Hal.Cell.Clamp.Finish THEN
           #Device.Processed := FALSE;
           IF #Unit.CarrierIndex = 0 THEN
               #Device.Processed := TRUE;
           ELSE
               #Device.Processed := "FRK_PartProcessed"(Core := #Core, Unit := #Unit, Status := #Status, Part := #Part, AlarmLog := #AlarmLog, Verdict := #Hal.Cell.Clamp.Verdict, Reason := #Hal.Cell.Clamp.Diag.ReasonCode);
           END_IF;
           IF #Device.Processed THEN
               #Device.Cycles := #Device.Cycles + 1;
               IF #Unit.StopReq THEN
                   "FRK_Complete"(Core := #Core,
                                  Status := #Status);
               ELSE
                   #Device.Received := "FRK_PartReceived"(Core := #Core, Unit := #Unit, Status := #Status, Part := #Part, AlarmLog := #AlarmLog);
                   IF #Device.Received THEN
                       "FRK_PartStarted"(Unit := #Unit,
                                         Status := #Status,
                                         Part := #Part,
                                         AlarmLog := #AlarmLog);
                   END_IF;
               END_IF;
           END_IF;
       END_IF;
       // ---- GENERATED: end dispatch
   END_IF;
   "FRK_End"(Core := #Core,
             Status := #Status,
             Busy => #Busy,
             Done => #Done,
             Error => #Error,
             Aborted => #Aborted,
             Held => #Held,
             ErrorID => #ErrorID,
             Timing => #Timing);
   "FRK_DecisionCyclic"(Owner := #Core.RegIndex,
                        Busy := #Core.Exec = 1,
                        Reset := #Startup OR #Unit.EvReset OR #Core.EvModeChanged,
                        AlarmLog := #AlarmLog);
   "FRK_DecisionPublish"(Owner := #Core.RegIndex,
                         Decision := #Decision,
                         DecisionAnswer := #DecisionAnswer);
   IF NOT #Unit.EvReset THEN
       "FRK_AlarmCapture"(AlarmLog := #AlarmLog,
                          Core := #Core,
                          Status := #Status);
       "FRK_Capture_DeclarationCell"(Module := #Cell,
                                     AlarmLog := #AlarmLog);
       "FRK_AlarmEnd"(AlarmLog := #AlarmLog);
   END_IF;
   IF #Core.RegIndex > 0 THEN
       "FRK_Registry".Rows[#Core.RegIndex].AlarmBlocking := #AlarmLog.Blocking;
   END_IF;
   #Unit.AlarmBlocking := "FRK_AlarmTreeBlocking"(Owner := #Core.RegIndex);
   "FRK_AccessPersist"(Access := #Access,
                       Unit := #Unit,
                       Response := #HmiResponse,
                       SourcePath := STRING_TO_WSTRING(#Status.Name),
                       AlarmLog := #AlarmLog);
   "FRK_AccessFinish"(Access := #Access,
                      Unit := #Unit,
                      Response := #HmiResponse,
                      SourcePath := STRING_TO_WSTRING(#Status.Name),
                      AlarmLog := #AlarmLog,
                      Revision := #ConfigRev);
   "FRK_UnitFinish"(Core := #Core,
                    Unit := #Unit,
                    Response := #HmiResponse,
                    Status := #Status,
                    Part := #Part,
                    AlarmLog := #AlarmLog,
                    History := #History,
                    Head := #HistoryHead);
   #ModeActivePublished := #Unit.Mode;
   #RunningPublished := #Core.Exec = 1;
   #StopPendingPublished := #Unit.StopReq AND #Core.Exec = 1;
   #GoodCount := #Unit.Good;
   #NokCount := #Unit.Nok;
   #ReworkCount := #Unit.Rework;
   #NokReason := #Unit.NokReason;
   // ---- AUTHORED: unconditional cyclic/derived data
   #OutImm.Cycles := #Device.Cycles;
   #OutImm.ExitCalls := #Device.ExitCalls;
   #OutImm.Changes := #Device.Changes;
   #OutImm.Resets := #Device.Resets;
   #OutImm.AtHome := "FRK_State"(Idx := 1, Key := 'project.state.atHome', Ok := #Hal.Cell.Clamp.Sample = 0, Flags := #StateFlags, Count := #StateFlagCount, Touched := #StateTouched);
   // ---- GENERATED: frame end
END_FUNCTION_BLOCK

FUNCTION "FRK_AccessAudit" : Void   // FC53, SCL
{ S7_Optimized_Access := 'TRUE' }
VERSION : 0.1
// stored: AutoNumber true, IsIECCheckEnabled false, SetENOAutomatically false, UDAEnableTagReadback false
   VAR_INPUT
      What : WString;
      Who : String;
      SourcePath : WString;
   END_VAR
   VAR_IN_OUT
      AlarmLog : "FRK_AlarmLog";
   END_VAR
   VAR_TEMP
      Description : WString[480];
   END_VAR
BEGIN

   #Description := CONCAT(IN1 := #What, IN2 := WSTRING#': ');
   #Description := CONCAT(IN1 := #Description, IN2 := STRING_TO_WSTRING(#Who));
   "FRK_AlarmMessage"(AlarmLog := #AlarmLog,
                      Reason := 0,
                      Description := #Description,
                      SourcePath := #SourcePath);
END_FUNCTION

FUNCTION "FRK_AccessCancel" : Void   // FC48, SCL
{ S7_Optimized_Access := 'TRUE' }
VERSION : 0.1
// stored: AutoNumber true, IsIECCheckEnabled false, SetENOAutomatically false, UDAEnableTagReadback false
   VAR_IN_OUT
      Access : "FRK_Access";
   END_VAR
   VAR_TEMP
      Index : DInt;
   END_VAR
BEGIN

   #Access.LoginBusy := FALSE;
   #Access.CandidateUser := '';
   #Access.CandidateLevel := 0;
   #Access.Round := 0;
   FOR #Index := 0 TO 15 DO
       #Access.Salt[#Index] := 0;
   END_FOR;
   FOR #Index := 0 TO 31 DO
       #Access.Digest[#Index] := 0;
       #Access.Expected[#Index] := 0;
   END_FOR;
END_FUNCTION

FUNCTION "FRK_AccessCyclic" : Void   // FC54, SCL
{ S7_Optimized_Access := 'TRUE' }
VERSION : 0.1
// stored: AutoNumber true, IsIECCheckEnabled false, SetENOAutomatically false, UDAEnableTagReadback false
   VAR_INPUT
      Startup : Bool;
      SourcePath : WString;
   END_VAR
   VAR_IN_OUT
      Access : "FRK_Access";
      AlarmLog : "FRK_AlarmLog";
      Revision : UDInt;
   END_VAR
   VAR_TEMP
      Data : Array[0..47] of Byte;
      Index : DInt;
      Difference : Byte;
      HashOk : Bool;
   END_VAR
BEGIN

   #Access.LoginTimeoutMs := 6000;
   IF #Startup THEN
       "FRK_AccessLogout"(Access := #Access);
       #Access.LoginResultSequence := 0;
   END_IF;
   IF #Access.ProviderGeneration <> "FRK_LocalUsers".Generation OR NOT "FRK_AccessStorage".UsersReady THEN
       IF #Access.CurrentLevel > 0 THEN
           "FRK_AccessAudit"(AlarmLog := #AlarmLog,
                             What := WSTRING#'std.audit.autoLogout',
                             Who := #Access.CurrentUser,
                             SourcePath := #SourcePath);
           "FRK_AccessDropSession"(Access := #Access);
           #Revision := "FRK_ConfigRevision"(Previous := #Revision);
       END_IF;
       IF #Access.LoginBusy THEN
           #Access.CandidateLevel := 0;
       END_IF;
       #Access.ProviderGeneration := "FRK_LocalUsers".Generation;
   END_IF;
   IF #Access.CurrentLevel > 0 AND #Access.Policy.SessionTimeout > T#0ms THEN
       IF "FRK_Elapsed"(NewMs := "FRK_Clock".NowMs, OldMs := #Access.LastActivity) >= DINT_TO_UDINT(TIME_TO_DINT(#Access.Policy.SessionTimeout)) THEN
           "FRK_AccessAudit"(AlarmLog := #AlarmLog,
                             What := WSTRING#'std.audit.autoLogout',
                             Who := #Access.CurrentUser,
                             SourcePath := #SourcePath);
           // Expiring the old session does not discard a separately committed
           // credential attempt. Explicit logout cancels both.
           "FRK_AccessDropSession"(Access := #Access);
           #Revision := "FRK_ConfigRevision"(Previous := #Revision);
       END_IF;
   END_IF;
   IF NOT #Access.LoginBusy THEN
       RETURN;
   END_IF;
   // One compression per active scan; never run all PIN rounds in one scan.
   FOR #Index := 0 TO 31 DO
       #Data[#Index] := #Access.Digest[#Index];
   END_FOR;
   FOR #Index := 0 TO 15 DO
       #Data[32 + #Index] := #Access.Salt[#Index];
   END_FOR;
   #HashOk := "FRK_Sha256Pin"(Data := #Data, Size := 48, Digest := #Access.Digest);
   FOR #Index := 0 TO 47 DO
       #Data[#Index] := 0;
   END_FOR;
   #Access.Round := #Access.Round + 1;
   IF NOT #HashOk OR "FRK_Elapsed"(NewMs := "FRK_Clock".NowMs, OldMs := #Access.LoginSince) >= #Access.LoginTimeoutMs THEN
       #Access.CandidateLevel := 0;
   ELSIF #Access.Round < 256 THEN
       RETURN;
   END_IF;
   #Difference := 0;
   FOR #Index := 0 TO 31 DO
       #Difference := #Difference OR (#Access.Digest[#Index] XOR #Access.Expected[#Index]);
   END_FOR;
   #Access.LoginFailed := #Difference <> 0 OR #Access.CandidateLevel = 0 OR NOT #Access.ProviderEnabled OR NOT "FRK_AccessStorage".UsersReady OR #Access.CandidateGeneration <> "FRK_LocalUsers".Generation;
   IF #Access.LoginFailed THEN
       "FRK_AccessAudit"(AlarmLog := #AlarmLog,
                         What := WSTRING#'std.audit.loginFailed',
                         Who := #Access.CandidateUser,
                         SourcePath := #SourcePath);
   ELSE
       #Access.CurrentUser := #Access.CandidateUser;
       #Access.CurrentLevel := #Access.CandidateLevel;
       #Access.LastActivity := "FRK_Clock".NowMs;
       #Access.SessionGeneration := "FRK_AccessNext"(Previous := #Access.SessionGeneration);
       #Revision := "FRK_ConfigRevision"(Previous := #Revision);
       "FRK_AccessAudit"(AlarmLog := #AlarmLog,
                         What := WSTRING#'std.audit.login',
                         Who := #Access.CurrentUser,
                         SourcePath := #SourcePath);
   END_IF;
   #Access.LoginResultSequence := #Access.LoginSequence;
   "FRK_AccessCancel"(Access := #Access);
END_FUNCTION

FUNCTION "FRK_AccessDropSession" : Void   // FC50, SCL
{ S7_Optimized_Access := 'TRUE' }
VERSION : 0.1
// stored: AutoNumber true, IsIECCheckEnabled false, SetENOAutomatically false, UDAEnableTagReadback false
   VAR_IN_OUT
      Access : "FRK_Access";
   END_VAR
BEGIN

   #Access.CurrentLevel := 0;
   #Access.CurrentUser := '';
   #Access.LoginFailed := FALSE;
   #Access.SessionGeneration := "FRK_AccessNext"(Previous := #Access.SessionGeneration);
END_FUNCTION

FUNCTION "FRK_AccessFinish" : Void   // FC55, SCL
{ S7_Optimized_Access := 'TRUE' }
VERSION : 0.1
// stored: AutoNumber true, IsIECCheckEnabled false, SetENOAutomatically false, UDAEnableTagReadback false
   VAR_INPUT
      Unit : "FRK_Unit";
      Response : "ST_HmiResponse";
      SourcePath : WString;
   END_VAR
   VAR_IN_OUT
      Access : "FRK_Access";
      AlarmLog : "FRK_AlarmLog";
      Revision : UDInt;
   END_VAR
   VAR_TEMP
      What : WString[160];
      AuditPath : WString[255];
   END_VAR
BEGIN

   IF NOT #Unit.RequestPending THEN
       RETURN;
   END_IF;
   CASE #Unit.Request.Kind OF
       23, 15,
       16, 17,
       1:
           RETURN;
       2:
           "FRK_AccessAudit"(AlarmLog := #AlarmLog,
                             What := WSTRING#'std.audit.logout',
                             Who := #Unit.RequestUser,
                             SourcePath := #SourcePath);
           #Revision := "FRK_ConfigRevision"(Previous := #Revision);
           RETURN;
       ELSE
           #What := WSTRING#'std.audit.accessDenied';
   END_CASE;
   IF #Response.Accepted THEN
       #What := WSTRING#'std.audit.operatorAction';
       IF #Access.CurrentLevel > 0 THEN
           #Access.LastActivity := "FRK_Clock".NowMs;
       END_IF;
       IF #Unit.Request.Kind = 24 OR #Unit.Request.Kind = 25 THEN
           #Revision := "FRK_ConfigRevision"(Previous := #Revision);
       END_IF;
   END_IF;
   #AuditPath := #SourcePath;
   IF #Unit.Request.Kind = 11 THEN
       IF #Response.Accepted THEN
           #AuditPath := #Unit.Request.TargetPath;
       END_IF;
       IF #Response.Accepted THEN
           #What := WSTRING#'std.audit.manualCommandAccepted';
       ELSE
           #What := WSTRING#'std.audit.manualCommandRejected';
       END_IF;
   END_IF;
   #What := CONCAT(IN1 := #What, IN2 := WSTRING#' kind=');
   #What := CONCAT(IN1 := #What, IN2 := DINT_TO_WSTRING(#Unit.Request.Kind));
   #What := CONCAT(IN1 := #What, IN2 := WSTRING#' value=');
   #What := CONCAT(IN1 := #What, IN2 := DINT_TO_WSTRING(#Unit.Request.IntValue));
   "FRK_AccessAudit"(AlarmLog := #AlarmLog,
                     What := #What,
                     Who := #Unit.RequestUser,
                     SourcePath := #AuditPath);
END_FUNCTION

FUNCTION "FRK_AccessLogin" : Void   // FC52, SCL
{ S7_Optimized_Access := 'TRUE' }
VERSION : 0.1
// stored: AutoNumber true, IsIECCheckEnabled false, SetENOAutomatically false, UDAEnableTagReadback false
   VAR_INPUT
      User : String;
      Secret : String;
      Sequence : UDInt;
   END_VAR
   VAR_IN_OUT
      Access : "FRK_Access";
   END_VAR
   VAR_TEMP
      Data : Array[0..47] of Byte;
      Index : DInt;
      Slot : DInt;
      Size : Int;
      HashOk : Bool;
   END_VAR
BEGIN

   "FRK_AccessCancel"(Access := #Access);
   #Access.LoginFailed := FALSE;
   #Access.LoginSequence := #Sequence;
   #Access.CandidateGeneration := "FRK_LocalUsers".Generation;
   #Access.LoginSince := "FRK_Clock".NowMs;
   #Access.LoginTimeoutMs := 6000;
   #Access.CandidateUser := #User;
   // Unknown users execute the same bounded work with a dummy salt/digest.
   IF #Access.ProviderEnabled AND "FRK_AccessStorage".UsersReady AND "FRK_LocalUsers".Count >= 0 AND "FRK_LocalUsers".Count <= 16 THEN
       FOR #Slot := 1 TO "FRK_LocalUsers".Count DO
           IF #User <> '' AND "FRK_LocalUsers".Rows[#Slot].User = #User THEN
               IF "FRK_LocalUsers".Rows[#Slot].Level >= 1 AND "FRK_LocalUsers".Rows[#Slot].Level <= 4 THEN
                   #Access.CandidateLevel := "FRK_LocalUsers".Rows[#Slot].Level;
                   #Access.Salt := "FRK_LocalUsers".Rows[#Slot].Salt;
                   #Access.Expected := "FRK_LocalUsers".Rows[#Slot].PinHash;
               END_IF;
               EXIT;
           END_IF;
       END_FOR;
   END_IF;
   FOR #Index := 0 TO 47 DO
       #Data[#Index] := 0;
   END_FOR;
   FOR #Index := 0 TO 15 DO
       #Data[#Index] := #Access.Salt[#Index];
   END_FOR;
   #Size := LEN(#Secret);
   IF #Size > 32 THEN
       #Size := 0;
       #Access.CandidateLevel := 0;
   END_IF;
   FOR #Index := 1 TO #Size DO
       #Data[15 + #Index] := CHAR_TO_BYTE(#Secret[#Index]);
   END_FOR;
   #HashOk := "FRK_Sha256Pin"(Data := #Data, Size := 16 + INT_TO_DINT(#Size), Digest := #Access.Digest);
   FOR #Index := 0 TO 47 DO
       #Data[#Index] := 0;
   END_FOR;
   #Access.LoginBusy := #HashOk;
END_FUNCTION

FUNCTION "FRK_AccessLogout" : Void   // FC49, SCL
{ S7_Optimized_Access := 'TRUE' }
VERSION : 0.1
// stored: AutoNumber true, IsIECCheckEnabled false, SetENOAutomatically false, UDAEnableTagReadback false
   VAR_IN_OUT
      Access : "FRK_Access";
   END_VAR
BEGIN

   "FRK_AccessCancel"(Access := #Access);
   "FRK_AccessDropSession"(Access := #Access);
END_FUNCTION

FUNCTION "FRK_AccessNext" : UDInt   // FC51, SCL
{ S7_Optimized_Access := 'TRUE' }
VERSION : 0.1
// stored: AutoNumber true, IsIECCheckEnabled false, SetENOAutomatically false, UDAEnableTagReadback false
   VAR_INPUT
      Previous : UDInt;
   END_VAR
BEGIN

   IF #Previous = UDINT#4294967295 THEN
       #FRK_AccessNext := 1;
   ELSE
       #FRK_AccessNext := #Previous + 1;
   END_IF;
END_FUNCTION

FUNCTION "FRK_AccessPersist" : Void   // FC68, SCL
{ S7_Optimized_Access := 'TRUE' }
VERSION : 0.1
// stored: AutoNumber true, IsIECCheckEnabled false, SetENOAutomatically false, UDAEnableTagReadback false
   VAR_INPUT
      Unit : "FRK_Unit";
      SourcePath : WString;
   END_VAR
   VAR_IN_OUT
      Access : "FRK_Access";
      Response : "ST_HmiResponse";
      AlarmLog : "FRK_AlarmLog";
   END_VAR
   VAR_TEMP
      Diag : "ST_Diagnostic";
      Accepted : Bool;
   END_VAR
BEGIN

   IF #Unit.RequestPending AND #Unit.Request.Kind = 31 AND #Access.PolicyLost THEN
       // Explicit ENGINEER acknowledgement accepts the restrictive fallback.
       #Response.Accepted := #Access.CurrentLevel >= 3 AND #Access.PolicySlot > 0;
       IF #Response.Accepted THEN
           "FRK_AccessPolicySave"(Access := #Access,
                                  Scope := WSTRING_TO_STRING(#SourcePath));
           #Access.PolicyLost := FALSE;
           #Response.Diagnostic := WSTRING#'';
       ELSE
           #Response.Diagnostic := WSTRING#'std.error.configRestoreAckRefused';
       END_IF;
   ELSIF #Unit.RequestPending AND #Response.Accepted AND NOT #Access.PolicyLost AND (#Unit.Request.Kind = 24 OR #Unit.Request.Kind = 25) THEN
       "FRK_AccessPolicySave"(Access := #Access,
                              Scope := WSTRING_TO_STRING(#SourcePath));
   END_IF;
   IF #Access.PolicyLost AND #Access.PolicyLossAlarm = 0 THEN
       #Diag := "FRK_UnitScratch".EmptyDiagnostic;
       #Diag.ReasonCode := 2040;
       #Diag.Description := WSTRING#'std.error.configRestoreLost';
       #Diag.SourcePath := #SourcePath;
       #Access.PolicyLossAlarm := "FRK_AlarmRaise"(AlarmLog := #AlarmLog, Diag := #Diag, ResetClass := 0);
   ELSIF NOT #Access.PolicyLost AND #Access.PolicyLossAlarm > 0 THEN
       #Accepted := "FRK_AlarmGone"(AlarmLog := #AlarmLog, Slot := #Access.PolicyLossAlarm);
       #Access.PolicyLossAlarm := 0;
   END_IF;
   IF "FRK_AccessStorage".UsersLost AND #Access.PolicySlot > 0 AND #Access.UserLossAlarm = 0 THEN
       #Diag := "FRK_UnitScratch".EmptyDiagnostic;
       #Diag.ReasonCode := 2040;
       #Diag.Description := WSTRING#'std.error.accessRestoreLost';
       #Diag.SourcePath := #SourcePath;
       #Access.UserLossAlarm := "FRK_AlarmRaise"(AlarmLog := #AlarmLog, Diag := #Diag, ResetClass := 0);
   ELSIF NOT "FRK_AccessStorage".UsersLost AND #Access.UserLossAlarm > 0 THEN
       #Accepted := "FRK_AlarmGone"(AlarmLog := #AlarmLog, Slot := #Access.UserLossAlarm);
       #Access.UserLossAlarm := 0;
   END_IF;
END_FUNCTION

FUNCTION "FRK_AccessPolicyBoot" : Void   // FC67, SCL
{ S7_Optimized_Access := 'TRUE' }
VERSION : 0.1
// stored: AutoNumber true, IsIECCheckEnabled false, SetENOAutomatically false, UDAEnableTagReadback false
   VAR_INPUT
      Startup : Bool;
      Root : Bool;
      Scope : String;
   END_VAR
   VAR_IN_OUT
      Access : "FRK_Access";
   END_VAR
   VAR_TEMP
      Index : Int;
      FreeSlot : Int;
   END_VAR
BEGIN

   IF NOT #Startup THEN
       RETURN;
   END_IF;
   #Access.PolicySlot := 0;
   #Access.PolicyLost := FALSE;
   #Access.PolicyLossAlarm := 0;
   #Access.UserLossAlarm := 0;
   IF NOT #Root THEN
       RETURN;
   END_IF;
   #FreeSlot := 0;
   FOR #Index := 1 TO 2 DO
       IF "FRK_AccessPolicies".Rows[#Index].Scope = #Scope THEN
           IF #Access.PolicySlot <> 0 THEN
               #Access.PolicyLost := TRUE;
           ELSE
               #Access.PolicySlot := #Index;
           END_IF;
       ELSIF #FreeSlot = 0 AND NOT "FRK_AccessPolicies".Rows[#Index].Initialized AND "FRK_AccessPolicies".Rows[#Index].Scope = '' AND "FRK_AccessPolicies".Rows[#Index].SchemaVersion = 0 AND "FRK_AccessPolicies".Rows[#Index].Generation = 0 AND "FRK_AccessPolicies".Rows[#Index].Checksum = DWORD#0 THEN
           #FreeSlot := #Index;
       END_IF;
   END_FOR;
   IF #Access.PolicySlot > 0 THEN
       IF NOT #Access.PolicyLost AND "FRK_AccessPolicyValid"(Image := "FRK_AccessPolicies".Rows[#Access.PolicySlot]) THEN
           #Access.Policy := "FRK_AccessPolicies".Rows[#Access.PolicySlot].Policy;
       ELSE
           #Access.PolicyLost := TRUE;
       END_IF;
   ELSIF #FreeSlot > 0 THEN
       #Access.PolicySlot := #FreeSlot;
       "FRK_AccessPolicySave"(Access := #Access,
                              Scope := #Scope);
   ELSE
       #Access.PolicyLost := TRUE;
   END_IF;
   IF #Access.PolicyLost THEN
       // Do not silently reopen actions after losing commissioned policy.
       #Access.Policy := "FRK_AccessStorage".EmptyPolicy;
       FOR #Index := 0 TO 11 DO
           #Access.Policy.Required[#Index] := 4;
       END_FOR;
   END_IF;
END_FUNCTION

FUNCTION "FRK_AccessPolicyCrc" : DWord   // FC63, SCL
{ S7_Optimized_Access := 'TRUE' }
VERSION : 0.1
// stored: AutoNumber true, IsIECCheckEnabled false, SetENOAutomatically false, UDAEnableTagReadback false
   VAR_IN_OUT
      Image : "FRK_AccessPolicyImage";
   END_VAR
   VAR_TEMP
      Work : DWord;
      Index : Int;
      Size : Int;
   END_VAR
BEGIN

   #Work := "FRK_CrcNumber"(Previous := DWORD#16#FFFFFFFF, Value := UINT_TO_UDINT(#Image.SchemaVersion));
   IF #Image.Initialized THEN
       #Work := "FRK_CrcByte"(Previous := #Work, Value := BYTE#1);
   ELSE
       #Work := "FRK_CrcByte"(Previous := #Work, Value := BYTE#0);
   END_IF;
   #Work := "FRK_CrcNumber"(Previous := #Work, Value := #Image.Generation);
   #Size := LEN(#Image.Scope);
   #Work := "FRK_CrcNumber"(Previous := #Work, Value := INT_TO_UDINT(#Size));
   FOR #Index := 1 TO #Size DO
       #Work := "FRK_CrcByte"(Previous := #Work, Value := CHAR_TO_BYTE(#Image.Scope[#Index]));
   END_FOR;
   FOR #Index := 0 TO 11 DO
       #Work := "FRK_CrcNumber"(Previous := #Work, Value := DINT_TO_UDINT(#Image.Policy.Required[#Index]));
   END_FOR;
   #Work := "FRK_CrcNumber"(Previous := #Work, Value := DINT_TO_UDINT(TIME_TO_DINT(#Image.Policy.SessionTimeout)));
   #FRK_AccessPolicyCrc := NOT #Work;
END_FUNCTION

FUNCTION "FRK_AccessPolicySave" : Void   // FC66, SCL
{ S7_Optimized_Access := 'TRUE' }
VERSION : 0.1
// stored: AutoNumber true, IsIECCheckEnabled false, SetENOAutomatically false, UDAEnableTagReadback false
   VAR_INPUT
      Scope : String;
   END_VAR
   VAR_IN_OUT
      Access : "FRK_Access";
   END_VAR
BEGIN

   IF #Access.PolicySlot < 1 OR #Access.PolicySlot > 2 THEN
       RETURN;
   END_IF;
   IF #Scope = '' OR NOT "FRK_AccessPolicyShape"(Policy := #Access.Policy) THEN
       #Access.PolicyLost := TRUE;
       RETURN;
   END_IF;
   "FRK_AccessPolicies".Rows[#Access.PolicySlot].SchemaVersion := 1;
   "FRK_AccessPolicies".Rows[#Access.PolicySlot].Initialized := TRUE;
   "FRK_AccessPolicies".Rows[#Access.PolicySlot].Scope := #Scope;
   "FRK_AccessPolicies".Rows[#Access.PolicySlot].Generation := "FRK_AccessNext"(Previous := "FRK_AccessPolicies".Rows[#Access.PolicySlot].Generation);
   "FRK_AccessPolicies".Rows[#Access.PolicySlot].Policy := #Access.Policy;
   "FRK_AccessPolicies".Rows[#Access.PolicySlot].Checksum := "FRK_AccessPolicyCrc"(Image := "FRK_AccessPolicies".Rows[#Access.PolicySlot]);
END_FUNCTION

FUNCTION "FRK_AccessPolicyShape" : Bool   // FC64, SCL
{ S7_Optimized_Access := 'TRUE' }
VERSION : 0.1
// stored: AutoNumber true, IsIECCheckEnabled false, SetENOAutomatically false, UDAEnableTagReadback false
   VAR_IN_OUT
      Policy : "ST_AccessPolicy";
   END_VAR
   VAR_TEMP
      Index : Int;
   END_VAR
BEGIN

   #FRK_AccessPolicyShape := FALSE;
   IF #Policy.SessionTimeout < T#0ms OR #Policy.SessionTimeout > T#604800000ms THEN
       RETURN;
   END_IF;
   FOR #Index := 0 TO 11 DO
       IF #Policy.Required[#Index] < 0 OR #Policy.Required[#Index] > 4 THEN
           RETURN;
       END_IF;
   END_FOR;
   #FRK_AccessPolicyShape := TRUE;
END_FUNCTION

FUNCTION "FRK_AccessPolicyValid" : Bool   // FC65, SCL
{ S7_Optimized_Access := 'TRUE' }
VERSION : 0.1
// stored: AutoNumber true, IsIECCheckEnabled false, SetENOAutomatically false, UDAEnableTagReadback false
   VAR_IN_OUT
      Image : "FRK_AccessPolicyImage";
   END_VAR
   VAR_TEMP
      Index : Int;
   END_VAR
BEGIN

   #FRK_AccessPolicyValid := FALSE;
   IF NOT #Image.Initialized OR #Image.SchemaVersion <> 1 OR #Image.Scope = '' OR #Image.Generation = 0 OR NOT "FRK_AccessPolicyShape"(Policy := #Image.Policy) THEN
       RETURN;
   END_IF;
   #FRK_AccessPolicyValid := #Image.Checksum = "FRK_AccessPolicyCrc"(Image := #Image);
END_FUNCTION

FUNCTION "FRK_AccessRegisterHash" : Bool   // FC61, SCL
{ S7_Optimized_Access := 'TRUE' }
VERSION : 0.1
// stored: AutoNumber true, IsIECCheckEnabled false, SetENOAutomatically false, UDAEnableTagReadback false
   VAR_INPUT
      Record : "ST_UserRecord";
   END_VAR
   VAR_TEMP
      Slot : Int;
      Index : Int;
   END_VAR
BEGIN

   // Trusted composition/provider seam, never a remote credential editor.
   #FRK_AccessRegisterHash := FALSE;
   IF NOT "FRK_AccessStorage".UsersReady OR #Record.User = '' OR #Record.Level < 0 OR #Record.Level > 4 THEN
       RETURN;
   END_IF;
   #Slot := 0;
   FOR #Index := 1 TO DINT_TO_INT("FRK_LocalUsers".Count) DO
       IF "FRK_LocalUsers".Rows[#Index].User = #Record.User THEN
           #Slot := #Index;
           EXIT;
       END_IF;
   END_FOR;
   IF #Slot = 0 THEN
       IF "FRK_LocalUsers".Count = 16 THEN
           RETURN;
       END_IF;
       "FRK_LocalUsers".Count := "FRK_LocalUsers".Count + 1;
       #Slot := DINT_TO_INT("FRK_LocalUsers".Count);
   END_IF;
   "FRK_LocalUsers".Rows[#Slot] := #Record;
   #FRK_AccessRegisterHash := "FRK_AccessUsersCommit"();
END_FUNCTION

FUNCTION "FRK_AccessStoreBoot" : Void   // FC62, SCL
{ S7_Optimized_Access := 'TRUE' }
VERSION : 0.1
// stored: AutoNumber true, IsIECCheckEnabled false, SetENOAutomatically false, UDAEnableTagReadback false
   VAR_INPUT
      Startup : Bool;
   END_VAR
   VAR_TEMP
      Accepted : Bool;
   END_VAR
BEGIN

   IF NOT #Startup THEN
       RETURN;
   END_IF;
   "FRK_AccessStorage".UsersReady := FALSE;
   "FRK_AccessStorage".UsersLost := FALSE;
   // A virgin image may accept deliberate composition-root provisioning.
   IF NOT "FRK_AccessStorage".UsersCommissioned AND "FRK_LocalUsers".SchemaVersion = 0 AND "FRK_LocalUsers".Generation = 0 AND "FRK_LocalUsers".Checksum = DWORD#0 THEN
       #Accepted := "FRK_AccessUsersCommit"();
       "FRK_AccessStorage".UsersLost := NOT #Accepted;
   ELSIF "FRK_AccessStorage".UsersCommissioned AND "FRK_LocalUsers".SchemaVersion = 1 AND "FRK_LocalUsers".Generation > 0 AND "FRK_AccessUsersShape"() THEN
       "FRK_AccessStorage".UsersReady := "FRK_LocalUsers".Checksum = "FRK_AccessUsersCrc"();
       "FRK_AccessStorage".UsersLost := NOT "FRK_AccessStorage".UsersReady;
   ELSE
       "FRK_AccessStorage".UsersLost := TRUE;
   END_IF;
END_FUNCTION

FUNCTION "FRK_AccessUsersCommit" : Bool   // FC60, SCL
{ S7_Optimized_Access := 'TRUE' }
VERSION : 0.1
// stored: AutoNumber true, IsIECCheckEnabled false, SetENOAutomatically false, UDAEnableTagReadback false
BEGIN

   #FRK_AccessUsersCommit := "FRK_AccessUsersShape"();
   IF NOT #FRK_AccessUsersCommit THEN
       RETURN;
   END_IF;
   "FRK_LocalUsers".SchemaVersion := 1;
   "FRK_LocalUsers".Generation := "FRK_AccessNext"(Previous := "FRK_LocalUsers".Generation);
   "FRK_LocalUsers".Checksum := "FRK_AccessUsersCrc"();
   "FRK_AccessStorage".UsersCommissioned := TRUE;
   "FRK_AccessStorage".UsersReady := TRUE;
   "FRK_AccessStorage".UsersLost := FALSE;
END_FUNCTION

FUNCTION "FRK_AccessUsersCrc" : DWord   // FC58, SCL
{ S7_Optimized_Access := 'TRUE' }
VERSION : 0.1
// stored: AutoNumber true, IsIECCheckEnabled false, SetENOAutomatically false, UDAEnableTagReadback false
   VAR_TEMP
      Work : DWord;
      Slot : Int;
      Index : Int;
      Size : Int;
   END_VAR
BEGIN

   #Work := "FRK_CrcNumber"(Previous := DWORD#16#FFFFFFFF, Value := UINT_TO_UDINT("FRK_LocalUsers".SchemaVersion));
   #Work := "FRK_CrcNumber"(Previous := #Work, Value := "FRK_LocalUsers".Generation);
   #Work := "FRK_CrcNumber"(Previous := #Work, Value := DINT_TO_UDINT("FRK_LocalUsers".Count));
   // Unused rows are included: an altered dormant credential is not ignored.
   FOR #Slot := 1 TO 16 DO
       #Size := LEN("FRK_LocalUsers".Rows[#Slot].User);
       #Work := "FRK_CrcNumber"(Previous := #Work, Value := INT_TO_UDINT(#Size));
       FOR #Index := 1 TO #Size DO
           #Work := "FRK_CrcByte"(Previous := #Work, Value := CHAR_TO_BYTE("FRK_LocalUsers".Rows[#Slot].User[#Index]));
       END_FOR;
       #Work := "FRK_CrcNumber"(Previous := #Work, Value := DINT_TO_UDINT("FRK_LocalUsers".Rows[#Slot].Level));
       FOR #Index := 0 TO 15 DO
           #Work := "FRK_CrcByte"(Previous := #Work, Value := "FRK_LocalUsers".Rows[#Slot].Salt[#Index]);
       END_FOR;
       FOR #Index := 0 TO 31 DO
           #Work := "FRK_CrcByte"(Previous := #Work, Value := "FRK_LocalUsers".Rows[#Slot].PinHash[#Index]);
       END_FOR;
   END_FOR;
   #FRK_AccessUsersCrc := NOT #Work;
END_FUNCTION

FUNCTION "FRK_AccessUsersShape" : Bool   // FC59, SCL
{ S7_Optimized_Access := 'TRUE' }
VERSION : 0.1
// stored: AutoNumber true, IsIECCheckEnabled false, SetENOAutomatically false, UDAEnableTagReadback false
   VAR_TEMP
      Slot : Int;
      Other : Int;
   END_VAR
BEGIN

   #FRK_AccessUsersShape := FALSE;
   IF "FRK_LocalUsers".Count < 0 OR "FRK_LocalUsers".Count > 16 THEN
       RETURN;
   END_IF;
   FOR #Slot := 1 TO DINT_TO_INT("FRK_LocalUsers".Count) DO
       IF "FRK_LocalUsers".Rows[#Slot].User = '' OR "FRK_LocalUsers".Rows[#Slot].Level < 0 OR "FRK_LocalUsers".Rows[#Slot].Level > 4 THEN
           RETURN;
       END_IF;
       FOR #Other := 1 TO #Slot - 1 DO
           IF "FRK_LocalUsers".Rows[#Slot].User = "FRK_LocalUsers".Rows[#Other].User THEN
               RETURN;
           END_IF;
       END_FOR;
   END_FOR;
   #FRK_AccessUsersShape := TRUE;
END_FUNCTION

FUNCTION "FRK_AdoptFault" : Void   // FC10, SCL
{ S7_Optimized_Access := 'TRUE' }
VERSION : 0.1
// stored: AutoNumber true, IsIECCheckEnabled false, SetENOAutomatically false, UDAEnableTagReadback false
   VAR_INPUT
      Diag : "ST_Diagnostic";
   END_VAR
   VAR_IN_OUT
      Core : "FRK_Core";
      Status : "ST_ModuleStatus";
   END_VAR
BEGIN

   IF #Core.Exec = 3 THEN
       RETURN;
   END_IF;
   #Status.Diagnostic := #Diag;
   #Core.Exec := 3;
   #Core.Step := 0;
   #Core.Dispatch := FALSE;
   #Core.DiagTouched := TRUE;
END_FUNCTION

FUNCTION "FRK_AlarmBegin" : Void   // FC31, SCL
{ S7_Optimized_Access := 'TRUE' }
VERSION : 0.1
// stored: AutoNumber true, IsIECCheckEnabled false, SetENOAutomatically false, UDAEnableTagReadback false
   VAR_INPUT
      Startup : Bool;
   END_VAR
   VAR_IN_OUT
      AlarmLog : "FRK_AlarmLog";
   END_VAR
   VAR_TEMP
      Index : Int;
   END_VAR
BEGIN

   FOR #Index := 1 TO 16 DO
       #AlarmLog.Touched[#Index] := FALSE;
       IF #Startup THEN
           #AlarmLog.Active[#Index] := "FRK_UnitScratch".EmptyEvent;
           #AlarmLog.Automatic[#Index] := FALSE;
           #AlarmLog.ComeMs[#Index] := 0;
       END_IF;
   END_FOR;
   IF #Startup THEN
       FOR #Index := 1 TO 64 DO
           #AlarmLog.Ring[#Index] := "FRK_UnitScratch".EmptyEvent;
       END_FOR;
       #AlarmLog.RingHead := 0;
       #AlarmLog.RingUsed := 0;
       #AlarmLog.Truncated := FALSE;
   END_IF;
   IF #Startup AND #AlarmLog.HistorySlot > 0 THEN "FRK_AlarmHistoryClear"(AlarmLog := #AlarmLog);
   END_IF;
   "FRK_AlarmRefresh"(AlarmLog := #AlarmLog);
END_FUNCTION

FUNCTION "FRK_AlarmCapture" : Void   // FC37, SCL
{ S7_Optimized_Access := 'TRUE' }
VERSION : 0.1
// stored: AutoNumber true, IsIECCheckEnabled false, SetENOAutomatically false, UDAEnableTagReadback false
   VAR_IN_OUT
      AlarmLog : "FRK_AlarmLog";
      Core : "FRK_Core";
      Status : "ST_ModuleStatus";
   END_VAR
   VAR_TEMP
      Slot : Int;
   END_VAR
BEGIN

   #Slot := #Core.FaultSlot;
   IF #Slot < 1 OR #Slot > 16 THEN
       #Slot := 0;
   ELSIF NOT #AlarmLog.Automatic[#Slot] OR #AlarmLog.Active[#Slot].State <> 1
       OR #AlarmLog.Active[#Slot].SourcePath <> #Status.Diagnostic.SourcePath
       OR #AlarmLog.Active[#Slot].ReasonCode <> #Status.Diagnostic.ReasonCode
       OR #AlarmLog.Active[#Slot].Description <> #Status.Diagnostic.Description THEN
       #Slot := 0;
   END_IF;
   IF #Core.Exec = 3 AND NOT #Core.FaultHandled THEN
       IF #Slot = 0 THEN
           // Adopted first-outs share one active occurrence within this log.
           FOR #Slot := 1 TO 16 DO
               IF #AlarmLog.Automatic[#Slot] AND #AlarmLog.Active[#Slot].State = 1
                   AND #AlarmLog.Active[#Slot].SourcePath = #Status.Diagnostic.SourcePath
                   AND #AlarmLog.Active[#Slot].ReasonCode = #Status.Diagnostic.ReasonCode
                   AND #AlarmLog.Active[#Slot].Description = #Status.Diagnostic.Description THEN
                   EXIT;
               END_IF;
           END_FOR;
           IF #Slot > 16 THEN
               #Slot := "FRK_AlarmRaise"(AlarmLog := #AlarmLog, Diag := #Status.Diagnostic, ResetClass := 1);
           END_IF;
       END_IF;
       IF #Slot > 0 THEN
           #AlarmLog.Automatic[#Slot] := TRUE;
           #AlarmLog.Touched[#Slot] := TRUE;
       END_IF;
       #Core.FaultSlot := #Slot;
   ELSE
       #Core.FaultSlot := 0;
   END_IF;
END_FUNCTION

FUNCTION "FRK_AlarmClose" : Void   // FC33, SCL
{ S7_Optimized_Access := 'TRUE' }
VERSION : 0.1
// stored: AutoNumber true, IsIECCheckEnabled false, SetENOAutomatically false, UDAEnableTagReadback false
   VAR_INPUT
      Slot : Int;
   END_VAR
   VAR_IN_OUT
      AlarmLog : "FRK_AlarmLog";
   END_VAR
BEGIN

   IF #Slot < 1 OR #Slot > 16 THEN
       RETURN;
   END_IF;
   IF #AlarmLog.Active[#Slot].State = 0 THEN
       RETURN;
   END_IF;
   #AlarmLog.Active[#Slot].State := 0;
   IF #AlarmLog.RingHead < 0 OR #AlarmLog.RingHead > 64 THEN
       #AlarmLog.RingHead := 0;
   END_IF;
   #AlarmLog.RingHead := (#AlarmLog.RingHead MOD 64) + 1;
   IF #AlarmLog.RingUsed >= 64 THEN
       #AlarmLog.Truncated := TRUE;
   ELSE
       #AlarmLog.RingUsed := #AlarmLog.RingUsed + 1;
   END_IF;
   #AlarmLog.Ring[#AlarmLog.RingHead] := #AlarmLog.Active[#Slot];
   "FRK_AlarmHistoryAppend"(AlarmLog := #AlarmLog);
   #AlarmLog.Automatic[#Slot] := FALSE;
   "FRK_AlarmRefresh"(AlarmLog := #AlarmLog);
   "FRK_AlarmNotify"(AlarmLog := #AlarmLog,
                     Ev := #AlarmLog.Ring[#AlarmLog.RingHead]);
END_FUNCTION

FUNCTION "FRK_AlarmEnd" : Void   // FC38, SCL
{ S7_Optimized_Access := 'TRUE' }
VERSION : 0.1
// stored: AutoNumber true, IsIECCheckEnabled false, SetENOAutomatically false, UDAEnableTagReadback false
   VAR_IN_OUT
      AlarmLog : "FRK_AlarmLog";
   END_VAR
   VAR_TEMP
      Slot : Int;
      Gone : Bool;
   END_VAR
BEGIN

   FOR #Slot := 1 TO 16 DO
       IF #AlarmLog.Automatic[#Slot] AND NOT #AlarmLog.Touched[#Slot] THEN
           #Gone := "FRK_AlarmGone"(AlarmLog := #AlarmLog, Slot := #Slot);
       END_IF;
   END_FOR;
END_FUNCTION

FUNCTION "FRK_AlarmEventCrc" : DWord   // FC41, SCL
{ S7_Optimized_Access := 'TRUE' }
VERSION : 0.1
// stored: AutoNumber true, IsIECCheckEnabled false, SetENOAutomatically false, UDAEnableTagReadback false
   VAR_INPUT
      Ev : "ST_AlarmEvent";
   END_VAR
   VAR_TEMP
      Work : DWord;
      Index : Int;
      Size : Int;
      Code : Word;
      Wide : LWord;
   END_VAR
BEGIN

   #Work := DWORD#16#FFFFFFFF;
   #Work := "FRK_CrcNumber"(Previous := #Work,
                            Value := DINT_TO_UDINT(#Ev.ReasonCode));
   #Size := LEN(#Ev.Description);
   #Work := "FRK_CrcNumber"(Previous := #Work,
                            Value := INT_TO_UDINT(#Size));
   FOR #Index := 1 TO #Size DO
       #Code := WCHAR_TO_WORD(#Ev.Description[#Index]);
       #Work := "FRK_CrcByte"(Previous := #Work,
                              Value := WORD_TO_BYTE(#Code));
       #Work := "FRK_CrcByte"(Previous := #Work,
                              Value := WORD_TO_BYTE(SHR(IN := #Code, N := 8)));
   END_FOR;
   #Size := LEN(#Ev.SourcePath);
   #Work := "FRK_CrcNumber"(Previous := #Work,
                            Value := INT_TO_UDINT(#Size));
   FOR #Index := 1 TO #Size DO
       #Code := WCHAR_TO_WORD(#Ev.SourcePath[#Index]);
       #Work := "FRK_CrcByte"(Previous := #Work,
                              Value := WORD_TO_BYTE(#Code));
       #Work := "FRK_CrcByte"(Previous := #Work,
                              Value := WORD_TO_BYTE(SHR(IN := #Code, N := 8)));
   END_FOR;
   #Size := LEN(#Ev.IoTag);
   #Work := "FRK_CrcNumber"(Previous := #Work,
                            Value := INT_TO_UDINT(#Size));
   FOR #Index := 1 TO #Size DO
       #Work := "FRK_CrcByte"(Previous := #Work,
                              Value := CHAR_TO_BYTE(#Ev.IoTag[#Index]));
   END_FOR;
   #Size := LEN(#Ev.IoAddress);
   #Work := "FRK_CrcNumber"(Previous := #Work,
                            Value := INT_TO_UDINT(#Size));
   FOR #Index := 1 TO #Size DO
       #Work := "FRK_CrcByte"(Previous := #Work,
                              Value := CHAR_TO_BYTE(#Ev.IoAddress[#Index]));
   END_FOR;
   #Work := "FRK_CrcNumber"(Previous := #Work,
                            Value := DINT_TO_UDINT(#Ev.Severity));
   #Work := "FRK_CrcNumber"(Previous := #Work,
                            Value := DINT_TO_UDINT(#Ev.Category));
   #Work := "FRK_CrcNumber"(Previous := #Work,
                            Value := DINT_TO_UDINT(#Ev.ResetClass));
   #Work := "FRK_CrcNumber"(Previous := #Work,
                            Value := DINT_TO_UDINT(#Ev.State));
   #Wide := LINT_TO_LWORD(LDT_TO_LINT(#Ev.ComeAt));
   #Work := "FRK_CrcNumber"(Previous := #Work,
                            Value := DWORD_TO_UDINT(LWORD_TO_DWORD(#Wide)));
   #Work := "FRK_CrcNumber"(Previous := #Work,
                            Value := DWORD_TO_UDINT(LWORD_TO_DWORD(SHR(IN := #Wide, N := 32))));
   #Wide := LINT_TO_LWORD(LDT_TO_LINT(#Ev.GoneAt));
   #Work := "FRK_CrcNumber"(Previous := #Work,
                            Value := DWORD_TO_UDINT(LWORD_TO_DWORD(#Wide)));
   #Work := "FRK_CrcNumber"(Previous := #Work,
                            Value := DWORD_TO_UDINT(LWORD_TO_DWORD(SHR(IN := #Wide, N := 32))));
   #Wide := LINT_TO_LWORD(LDT_TO_LINT(#Ev.ResetAt));
   #Work := "FRK_CrcNumber"(Previous := #Work,
                            Value := DWORD_TO_UDINT(LWORD_TO_DWORD(#Wide)));
   #Work := "FRK_CrcNumber"(Previous := #Work,
                            Value := DWORD_TO_UDINT(LWORD_TO_DWORD(SHR(IN := #Wide, N := 32))));
   #Work := "FRK_CrcNumber"(Previous := #Work,
                            Value := DINT_TO_UDINT(TIME_TO_DINT(#Ev.Duration)));
   #Work := "FRK_CrcNumber"(Previous := #Work,
                            Value := BOOL_TO_UDINT(#Ev.Shelved));
   #Wide := LINT_TO_LWORD(LDT_TO_LINT(#Ev.ShelvedUntil));
   #Work := "FRK_CrcNumber"(Previous := #Work,
                            Value := DWORD_TO_UDINT(LWORD_TO_DWORD(#Wide)));
   #Work := "FRK_CrcNumber"(Previous := #Work,
                            Value := DWORD_TO_UDINT(LWORD_TO_DWORD(SHR(IN := #Wide, N := 32))));
   #Work := "FRK_CrcNumber"(Previous := #Work,
                            Value := BOOL_TO_UDINT(#Ev.ComeTimeSynchronized));
   #Work := "FRK_CrcNumber"(Previous := #Work,
                            Value := BOOL_TO_UDINT(#Ev.GoneTimeSynchronized));
   #Work := "FRK_CrcNumber"(Previous := #Work,
                            Value := BOOL_TO_UDINT(#Ev.ResetTimeSynchronized));
   #Work := "FRK_CrcNumber"(Previous := #Work,
                            Value := BOOL_TO_UDINT(#Ev.ShelfTimeSynchronized));
   #FRK_AlarmEventCrc := NOT #Work;
END_FUNCTION

FUNCTION "FRK_AlarmGone" : Bool   // FC34, SCL
{ S7_Optimized_Access := 'TRUE' }
VERSION : 0.1
// stored: AutoNumber true, IsIECCheckEnabled false, SetENOAutomatically false, UDAEnableTagReadback false
   VAR_INPUT
      Slot : Int;
   END_VAR
   VAR_IN_OUT
      AlarmLog : "FRK_AlarmLog";
   END_VAR
   VAR_TEMP
      Span : UDInt;
      Stamp : DTL;
      ResultCode : Int;
   END_VAR
BEGIN

   #FRK_AlarmGone := FALSE;
   IF #Slot < 1 OR #Slot > 16 THEN
       RETURN;
   END_IF;
   IF #AlarmLog.Active[#Slot].State <> 1 THEN
       RETURN;
   END_IF;
   #ResultCode := RD_SYS_T(OUT => #Stamp);
   IF #ResultCode = 0 THEN
       #AlarmLog.Active[#Slot].GoneAt := DTL_TO_LDT(#Stamp);
   END_IF;
   #AlarmLog.Active[#Slot].GoneTimeSynchronized := FALSE;
   #Span := "FRK_Elapsed"(NewMs := "FRK_Clock".NowMs, OldMs := #AlarmLog.ComeMs[#Slot]);
   IF #Span > 2147483647 THEN
       #Span := 2147483647;
   END_IF;
   #AlarmLog.Active[#Slot].Duration := DINT_TO_TIME(UDINT_TO_DINT(#Span));
   IF #AlarmLog.Active[#Slot].ResetClass = 0 THEN
       "FRK_AlarmClose"(AlarmLog := #AlarmLog,
                        Slot := #Slot);
   ELSE
       #AlarmLog.Active[#Slot].State := 2;
       #AlarmLog.Automatic[#Slot] := FALSE;
   END_IF;
   #FRK_AlarmGone := TRUE;
END_FUNCTION

FUNCTION "FRK_AlarmHistoryAppend" : Void   // FC45, SCL
{ S7_Optimized_Access := 'TRUE' }
VERSION : 0.1
// stored: AutoNumber true, IsIECCheckEnabled false, SetENOAutomatically false, UDAEnableTagReadback false
   VAR_IN_OUT
      AlarmLog : "FRK_AlarmLog";
   END_VAR
   VAR_TEMP
      Slot : Int;
      Head : Int;
   END_VAR
BEGIN

   #Slot := #AlarmLog.HistorySlot;
   #Head := #AlarmLog.RingHead;
   IF #Slot < 1 OR #Slot > 3 OR #Head < 1 OR #Head > 64 THEN
       RETURN;
   END_IF;
   "FRK_AlarmHistory".Rows[#Slot].Ring[#Head] := #AlarmLog.Ring[#Head];
   "FRK_AlarmHistory".Rows[#Slot].EventCrc[#Head] := "FRK_AlarmEventCrc"(Ev := #AlarmLog.Ring[#Head]);
   "FRK_AlarmHistoryHeaderSave"(AlarmLog := #AlarmLog);
END_FUNCTION

FUNCTION "FRK_AlarmHistoryBoot" : Void   // FC46, SCL
{ S7_Optimized_Access := 'TRUE' }
VERSION : 0.1
// stored: AutoNumber true, IsIECCheckEnabled false, SetENOAutomatically false, UDAEnableTagReadback false
   VAR_INPUT
      Startup : Bool;
      Scope : String;
   END_VAR
   VAR_IN_OUT
      AlarmLog : "FRK_AlarmLog";
   END_VAR
   VAR_TEMP
      Slot : Int;
      Index : Int;
      Used : Int;
      Head : Int;
      Valid : Bool;
   END_VAR
BEGIN

   IF NOT #Startup THEN
       RETURN;
   END_IF;
   #Slot := "FRK_AlarmHistoryIndex"(Scope := #Scope);
   #AlarmLog.HistorySlot := #Slot;
   IF #Slot < 1 OR #Slot > 3 THEN
       RETURN;
   END_IF;
   IF NOT "FRK_AlarmHistory".Commissioned[#Slot]
       AND "FRK_AlarmHistory".Rows[#Slot].SchemaVersion = 0
       AND "FRK_AlarmHistory".Rows[#Slot].Generation = 0
       AND "FRK_AlarmHistory".Rows[#Slot].Scope = ''
       AND "FRK_AlarmHistory".Rows[#Slot].Checksum = DWORD#0 THEN
       "FRK_AlarmHistory".Rows[#Slot].Scope := #Scope;
       "FRK_AlarmHistoryClear"(AlarmLog := #AlarmLog);
       RETURN;
   END_IF;
   #Used := "FRK_AlarmHistory".Rows[#Slot].RingUsed;
   #Head := "FRK_AlarmHistory".Rows[#Slot].RingHead;
   #Valid := "FRK_AlarmHistory".Rows[#Slot].SchemaVersion = 1
   AND "FRK_AlarmHistory".Rows[#Slot].Scope = #Scope
   AND "FRK_AlarmHistory".Rows[#Slot].Generation <> 0
   AND #Used >= 0 AND #Used <= 64
   AND #Head >= 0 AND #Head <= 64
   AND ((#Used = 0 AND #Head = 0) OR (#Used > 0 AND #Head > 0))
   AND (#Used = 64 OR #Head = #Used);
   IF #Valid THEN
       #Valid := "FRK_AlarmHistory".Rows[#Slot].Checksum = "FRK_AlarmHistoryHeaderCrc"(Slot := #Slot);
   END_IF;
   IF #Valid THEN
       FOR #Index := 1 TO #Used DO
           IF "FRK_AlarmHistory".Rows[#Slot].Ring[#Index].State <> 0
               OR "FRK_AlarmHistory".Rows[#Slot].Ring[#Index].ResetClass < 0
               OR "FRK_AlarmHistory".Rows[#Slot].Ring[#Index].ResetClass > 1
               OR "FRK_AlarmHistory".Rows[#Slot].Ring[#Index].Severity < 0
               OR "FRK_AlarmHistory".Rows[#Slot].Ring[#Index].Severity > 2
               OR "FRK_AlarmHistory".Rows[#Slot].Ring[#Index].Category < 0
               OR "FRK_AlarmHistory".Rows[#Slot].Ring[#Index].Category > 2
               OR "FRK_AlarmHistory".Rows[#Slot].Ring[#Index].SourcePath = WSTRING#''
               OR "FRK_AlarmHistory".Rows[#Slot].Ring[#Index].Description = WSTRING#''
               OR "FRK_AlarmHistory".Rows[#Slot].Ring[#Index].Duration < T#0ms
               OR "FRK_AlarmHistory".Rows[#Slot].EventCrc[#Index] <> "FRK_AlarmEventCrc"(Ev := "FRK_AlarmHistory".Rows[#Slot].Ring[#Index]) THEN
               #Valid := FALSE;
               EXIT;
           END_IF;
       END_FOR;
   END_IF;
   IF #Valid THEN
       FOR #Index := 1 TO #Used DO
           #AlarmLog.Ring[#Index] := "FRK_AlarmHistory".Rows[#Slot].Ring[#Index];
       END_FOR;
       #AlarmLog.RingHead := #Head;
       #AlarmLog.RingUsed := #Used;
       #AlarmLog.Truncated := "FRK_AlarmHistory".Rows[#Slot].Truncated;
   ELSE
       // Reject the whole image. The same public loss marker covers overflow
       // and rejected history; do not present a partial, apparently complete log.
       #AlarmLog.Truncated := TRUE;
       "FRK_AlarmHistory".Rows[#Slot].Scope := #Scope;
       "FRK_AlarmHistoryClear"(AlarmLog := #AlarmLog);
   END_IF;
END_FUNCTION

FUNCTION "FRK_AlarmHistoryClear" : Void   // FC44, SCL
{ S7_Optimized_Access := 'TRUE' }
VERSION : 0.1
// stored: AutoNumber true, IsIECCheckEnabled false, SetENOAutomatically false, UDAEnableTagReadback false
   VAR_IN_OUT
      AlarmLog : "FRK_AlarmLog";
   END_VAR
   VAR_TEMP
      Index : Int;
      Slot : Int;
   END_VAR
BEGIN

   #Slot := #AlarmLog.HistorySlot;
   IF #Slot < 1 OR #Slot > 3 THEN
       RETURN;
   END_IF;
   FOR #Index := 1 TO 64 DO
       "FRK_AlarmHistory".Rows[#Slot].Ring[#Index] := "FRK_UnitScratch".EmptyEvent;
       "FRK_AlarmHistory".Rows[#Slot].EventCrc[#Index] := DWORD#0;
   END_FOR;
   "FRK_AlarmHistoryHeaderSave"(AlarmLog := #AlarmLog);
END_FUNCTION

FUNCTION "FRK_AlarmHistoryHeaderCrc" : DWord   // FC42, SCL
{ S7_Optimized_Access := 'TRUE' }
VERSION : 0.1
// stored: AutoNumber true, IsIECCheckEnabled false, SetENOAutomatically false, UDAEnableTagReadback false
   VAR_INPUT
      Slot : Int;
   END_VAR
   VAR_TEMP
      Work : DWord;
      Index : Int;
      Size : Int;
   END_VAR
BEGIN

   #FRK_AlarmHistoryHeaderCrc := DWORD#0;
   IF #Slot < 1 OR #Slot > 3 THEN
       RETURN;
   END_IF;
   #Work := "FRK_CrcNumber"(Previous := DWORD#16#FFFFFFFF,
                            Value := UINT_TO_UDINT("FRK_AlarmHistory".Rows[#Slot].SchemaVersion));
   #Size := LEN("FRK_AlarmHistory".Rows[#Slot].Scope);
   #Work := "FRK_CrcNumber"(Previous := #Work,
                            Value := INT_TO_UDINT(#Size));
   FOR #Index := 1 TO #Size DO
       #Work := "FRK_CrcByte"(Previous := #Work,
                              Value := CHAR_TO_BYTE("FRK_AlarmHistory".Rows[#Slot].Scope[#Index]));
   END_FOR;
   #Work := "FRK_CrcNumber"(Previous := #Work,
                            Value := "FRK_AlarmHistory".Rows[#Slot].Generation);
   #Work := "FRK_CrcNumber"(Previous := #Work,
                            Value := INT_TO_UDINT("FRK_AlarmHistory".Rows[#Slot].RingHead));
   #Work := "FRK_CrcNumber"(Previous := #Work,
                            Value := INT_TO_UDINT("FRK_AlarmHistory".Rows[#Slot].RingUsed));
   #Work := "FRK_CrcNumber"(Previous := #Work,
                            Value := BOOL_TO_UDINT("FRK_AlarmHistory".Rows[#Slot].Truncated));
   FOR #Index := 1 TO 64 DO
       #Work := "FRK_CrcNumber"(Previous := #Work,
                                Value := DWORD_TO_UDINT("FRK_AlarmHistory".Rows[#Slot].EventCrc[#Index]));
   END_FOR;
   #FRK_AlarmHistoryHeaderCrc := NOT #Work;
END_FUNCTION

FUNCTION "FRK_AlarmHistoryHeaderSave" : Void   // FC43, SCL
{ S7_Optimized_Access := 'TRUE' }
VERSION : 0.1
// stored: AutoNumber true, IsIECCheckEnabled false, SetENOAutomatically false, UDAEnableTagReadback false
   VAR_IN_OUT
      AlarmLog : "FRK_AlarmLog";
   END_VAR
   VAR_TEMP
      Slot : Int;
   END_VAR
BEGIN

   #Slot := #AlarmLog.HistorySlot;
   IF #Slot < 1 OR #Slot > 3 THEN
       RETURN;
   END_IF;
   "FRK_AlarmHistory".Rows[#Slot].SchemaVersion := 1;
   "FRK_AlarmHistory".Rows[#Slot].Generation := "FRK_AccessNext"(Previous := "FRK_AlarmHistory".Rows[#Slot].Generation);
   "FRK_AlarmHistory".Rows[#Slot].RingHead := #AlarmLog.RingHead;
   "FRK_AlarmHistory".Rows[#Slot].RingUsed := #AlarmLog.RingUsed;
   "FRK_AlarmHistory".Rows[#Slot].Truncated := #AlarmLog.Truncated;
   "FRK_AlarmHistory".Rows[#Slot].Checksum := "FRK_AlarmHistoryHeaderCrc"(Slot := #Slot);
   "FRK_AlarmHistory".Commissioned[#Slot] := TRUE;
END_FUNCTION

FUNCTION "FRK_AlarmHistoryIndex" : Int   // FC40, SCL
{ S7_Optimized_Access := 'TRUE' }
VERSION : 0.1
// Reference-1500 LOCAL_RETAIN: closed history only, keyed by actual Unit scope.
//  No active alarms, commands, sessions or monotonic clocks are restored.
// stored: AutoNumber true, IsIECCheckEnabled false, SetENOAutomatically false, UDAEnableTagReadback false
   VAR_INPUT
      Scope : String;
   END_VAR
BEGIN

   #FRK_AlarmHistoryIndex := 0;
   IF #Scope = 'StationA' THEN
       #FRK_AlarmHistoryIndex := 1;
       RETURN;
   END_IF;
   IF #Scope = 'StationA.Satellite' THEN
       #FRK_AlarmHistoryIndex := 2;
       RETURN;
   END_IF;
   IF #Scope = 'StationB' THEN
       #FRK_AlarmHistoryIndex := 3;
       RETURN;
   END_IF;
END_FUNCTION

FUNCTION "FRK_AlarmMessage" : Void   // FC36, SCL
{ S7_Optimized_Access := 'TRUE' }
VERSION : 0.1
// stored: AutoNumber true, IsIECCheckEnabled false, SetENOAutomatically false, UDAEnableTagReadback false
   VAR_INPUT
      Reason : DInt;
      Description : WString;
      SourcePath : WString;
   END_VAR
   VAR_IN_OUT
      AlarmLog : "FRK_AlarmLog";
   END_VAR
   VAR_TEMP
      Diag : "ST_Diagnostic";
      Slot : Int;
      Gone : Bool;
   END_VAR
BEGIN

   #Diag := "FRK_UnitScratch".EmptyDiagnostic;
   #Diag.ReasonCode := #Reason;
   #Diag.Description := #Description;
   #Diag.SourcePath := #SourcePath;
   #Diag.Severity := 0;
   #Diag.Category := 2;
   #Slot := "FRK_AlarmRaise"(AlarmLog := #AlarmLog, Diag := #Diag, ResetClass := 0);
   IF #Slot > 0 THEN
       #Gone := "FRK_AlarmGone"(AlarmLog := #AlarmLog, Slot := #Slot);
   END_IF;
END_FUNCTION

FUNCTION "FRK_AlarmNotify" : Void   // FC29, SCL
{ S7_Optimized_Access := 'TRUE' }
VERSION : 0.1
// Core 8.3: one owning active list / closed ring, with optional event callback.
// stored: AutoNumber true, IsIECCheckEnabled false, SetENOAutomatically false, UDAEnableTagReadback false
   VAR_INPUT
      Ev : "ST_AlarmEvent";
   END_VAR
   VAR_IN_OUT
      AlarmLog : "FRK_AlarmLog";
   END_VAR
BEGIN

   IF #AlarmLog.SinkEnabled THEN
       "F_TestEventSink"(Ev := #Ev);
   END_IF;
END_FUNCTION

FUNCTION "FRK_AlarmOperatorReset" : Void   // FC35, SCL
{ S7_Optimized_Access := 'TRUE' }
VERSION : 0.1
// stored: AutoNumber true, IsIECCheckEnabled false, SetENOAutomatically false, UDAEnableTagReadback false
   VAR_IN_OUT
      AlarmLog : "FRK_AlarmLog";
   END_VAR
   VAR_TEMP
      Slot : Int;
      Gone : Bool;
      Stamp : DTL;
      ResultCode : Int;
   END_VAR
BEGIN

   FOR #Slot := 1 TO 16 DO
       IF #AlarmLog.Active[#Slot].State <> 0 AND #AlarmLog.Active[#Slot].ResetClass = 1 THEN
           IF #AlarmLog.Active[#Slot].State = 1 THEN
               #Gone := "FRK_AlarmGone"(AlarmLog := #AlarmLog, Slot := #Slot);
           END_IF;
           #ResultCode := RD_SYS_T(OUT => #Stamp);
           IF #ResultCode = 0 THEN
               #AlarmLog.Active[#Slot].ResetAt := DTL_TO_LDT(#Stamp);
           END_IF;
           #AlarmLog.Active[#Slot].ResetTimeSynchronized := FALSE;
           "FRK_AlarmClose"(AlarmLog := #AlarmLog,
                            Slot := #Slot);
       END_IF;
   END_FOR;
END_FUNCTION

FUNCTION "FRK_AlarmRaise" : Int   // FC32, SCL
{ S7_Optimized_Access := 'TRUE' }
VERSION : 0.1
// stored: AutoNumber true, IsIECCheckEnabled false, SetENOAutomatically false, UDAEnableTagReadback false
   VAR_INPUT
      Diag : "ST_Diagnostic";
      ResetClass : DInt;
   END_VAR
   VAR_IN_OUT
      AlarmLog : "FRK_AlarmLog";
   END_VAR
   VAR_TEMP
      Slot : Int;
      Stamp : DTL;
      ResultCode : Int;
      Rational : "ST_Diagnostic";
   END_VAR
BEGIN

   #FRK_AlarmRaise := 0;
   IF #ResetClass < 0 OR #ResetClass > 1
       OR #Diag.Severity < 0 OR #Diag.Severity > 2
       OR #Diag.Category < 0 OR #Diag.Category > 2
       OR #Diag.SourcePath = WSTRING#'' OR #Diag.Description = WSTRING#'' THEN
       RETURN;
   END_IF;
   FOR #Slot := 1 TO 16 DO
       IF #AlarmLog.Active[#Slot].State = 0 THEN
           #Rational := #Diag;
           "FRK_Rationalize"(Diag := #Rational);
           #AlarmLog.Active[#Slot] := "FRK_UnitScratch".EmptyEvent;
           #AlarmLog.Active[#Slot].ReasonCode := #Rational.ReasonCode;
           #AlarmLog.Active[#Slot].Description := #Rational.Description;
           #AlarmLog.Active[#Slot].SourcePath := #Rational.SourcePath;
           #AlarmLog.Active[#Slot].IoTag := #Rational.IoTag;
           #AlarmLog.Active[#Slot].IoAddress := #Rational.IoAddress;
           #AlarmLog.Active[#Slot].Severity := #Rational.Severity;
           #AlarmLog.Active[#Slot].Category := #Rational.Category;
           #AlarmLog.Active[#Slot].ResetClass := #ResetClass;
           #AlarmLog.Active[#Slot].State := 1;
           #AlarmLog.ComeMs[#Slot] := "FRK_Clock".NowMs;
           #AlarmLog.Automatic[#Slot] := FALSE;
           #AlarmLog.Touched[#Slot] := FALSE;
           #ResultCode := RD_SYS_T(OUT => #Stamp);
           IF #ResultCode = 0 THEN
               #AlarmLog.Active[#Slot].ComeAt := DTL_TO_LDT(#Stamp);
           END_IF;
           // The UTC source has no proven synchronization witness yet.
           #AlarmLog.Active[#Slot].ComeTimeSynchronized := FALSE;
           "FRK_AlarmRefresh"(AlarmLog := #AlarmLog);
           "FRK_AlarmNotify"(AlarmLog := #AlarmLog,
                             Ev := #AlarmLog.Active[#Slot]);
           #FRK_AlarmRaise := #Slot;
           RETURN;
       END_IF;
   END_FOR;
   #AlarmLog.Truncated := TRUE;
   "FRK_AlarmHistoryHeaderSave"(AlarmLog := #AlarmLog);
END_FUNCTION

FUNCTION "FRK_AlarmRefresh" : Void   // FC30, SCL
{ S7_Optimized_Access := 'TRUE' }
VERSION : 0.1
// stored: AutoNumber true, IsIECCheckEnabled false, SetENOAutomatically false, UDAEnableTagReadback false
   VAR_IN_OUT
      AlarmLog : "FRK_AlarmLog";
   END_VAR
   VAR_TEMP
      Index : Int;
   END_VAR
BEGIN

   #AlarmLog.NActive := 0;
   #AlarmLog.Blocking := FALSE;
   FOR #Index := 1 TO 16 DO
       IF #AlarmLog.Active[#Index].State <> 0 THEN
           #AlarmLog.NActive := #AlarmLog.NActive + 1;
           IF #AlarmLog.Active[#Index].ResetClass = 1 THEN
               #AlarmLog.Blocking := TRUE;
           END_IF;
       END_IF;
   END_FOR;
END_FUNCTION

FUNCTION "FRK_AlarmTreeBlocking" : Bool   // FC39, SCL
{ S7_Optimized_Access := 'TRUE' }
VERSION : 0.1
// stored: AutoNumber true, IsIECCheckEnabled false, SetENOAutomatically false, UDAEnableTagReadback false
   VAR_INPUT
      Owner : DInt;
   END_VAR
   VAR_TEMP
      Index : DInt;
      Ancestor : DInt;
      Depth : DInt;
   END_VAR
BEGIN

   #FRK_AlarmTreeBlocking := TRUE;
   IF "FRK_Registry".Fault OR #Owner < 1 OR #Owner > "FRK_Registry".Count OR "FRK_Registry".Count > 32 THEN
       RETURN;
   END_IF;
   FOR #Index := 1 TO "FRK_Registry".Count DO
       IF "FRK_Registry".Rows[#Index].AlarmBlocking THEN
           #Ancestor := #Index;
           FOR #Depth := 1 TO 32 DO
               IF #Ancestor = #Owner THEN
                   RETURN;
               END_IF;
               IF #Ancestor = 0 THEN
                   EXIT;
               END_IF;
               IF #Ancestor < 1 OR #Ancestor > "FRK_Registry".Count THEN
                   RETURN;
               END_IF;
               #Ancestor := "FRK_Registry".Rows[#Ancestor].Parent;
           END_FOR;
           IF #Depth > 32 AND #Ancestor <> 0 THEN
               RETURN;
           END_IF;
       END_IF;
   END_FOR;
   #FRK_AlarmTreeBlocking := FALSE;
END_FUNCTION

FUNCTION "FRK_Begin" : Void   // FC16, SCL
{ S7_Optimized_Access := 'TRUE' }
VERSION : 0.1
// stored: AutoNumber true, IsIECCheckEnabled false, SetENOAutomatically false, UDAEnableTagReadback false
   VAR_INPUT
      Execute : Bool;
      Abort : Bool;
      Command : DInt;
   END_VAR
   VAR_IN_OUT
      Core : "FRK_Core";
      Status : "ST_ModuleStatus";
   END_VAR
BEGIN

   #Core.EvInit := NOT #Core.Initialized;
   #Core.Initialized := TRUE;
   #Core.EvCommandStart := FALSE;
   #Core.EvAbort := FALSE;
   #Core.EvAbortInError := FALSE;
   #Core.HoldReq := FALSE;
   #Core.DiagTouched := FALSE;
   #Core.FaultHandled := FALSE;
   #Core.HookResult := 0;
   IF NOT #Execute AND (#Core.Armed OR #Core.ReleasePending) AND (#Core.Exec = 2 OR #Core.Exec = 3 OR #Core.Exec = 4) THEN
       #Core.Exec := 0;
       #Core.Armed := FALSE;
       #Core.HoldReason := 0;
       "FRK_ClearDiag"(Status := #Status);
   END_IF;
   IF #Execute AND NOT #Core.ExecPrev AND (#Core.Exec = 0 OR (#Core.Exec = 3 AND NOT #Core.Armed)) THEN
       #Core.Exec := 1;
       #Core.Armed := TRUE;
       #Core.Command := #Command;
       #Core.Step := 10;
       #Core.StartMs := "FRK_Clock".NowMs;
       #Core.LastNowMs := "FRK_Clock".NowMs;
       #Core.ActiveMs := 0;
       #Core.TimeoutMs := 0;
       #Core.CommandLabel := '';
       #Core.TimingOpen := TRUE;
       #Core.Held := FALSE;
       #Core.HoldReason := 0;
       "FRK_ClearDiag"(Status := #Status);
       #Core.EvCommandStart := TRUE;
   END_IF;
   #Core.DeltaMs := "FRK_Elapsed"(NewMs := "FRK_Clock".NowMs, OldMs := #Core.LastNowMs);
   #Core.LastNowMs := "FRK_Clock".NowMs;
   #Core.ExecPrev := #Execute;
   #Core.Dispatch := #Core.Exec = 1;
END_FUNCTION

FUNCTION "FRK_Capture_DeclarationCell" : Void   // FC145, SCL
{ S7_Optimized_Access := 'TRUE' }
VERSION : 0.1
// stored: AutoNumber true, IsIECCheckEnabled false, SetENOAutomatically false, UDAEnableTagReadback false
   VAR_IN_OUT
      Module : "FB_DeclarationCell";
      AlarmLog : "FRK_AlarmLog";
   END_VAR
BEGIN

   "FRK_AlarmCapture"(AlarmLog := #AlarmLog,
                      Core := #Module.Core,
                      Status := #Module.Status);
   "FRK_Capture_DeclarationCylinder"(Module := #Module.Clamp,
                                     AlarmLog := #AlarmLog);
   "FRK_Capture_DeclarationCylinder"(Module := #Module.Gate,
                                     AlarmLog := #AlarmLog);
END_FUNCTION

FUNCTION "FRK_Capture_DeclarationCylinder" : Void   // FC137, SCL
{ S7_Optimized_Access := 'TRUE' }
VERSION : 0.1
// stored: AutoNumber true, IsIECCheckEnabled false, SetENOAutomatically false, UDAEnableTagReadback false
   VAR_IN_OUT
      Module : "FB_DeclarationCylinder";
      AlarmLog : "FRK_AlarmLog";
   END_VAR
BEGIN

   "FRK_AlarmCapture"(AlarmLog := #AlarmLog,
                      Core := #Module.Core,
                      Status := #Module.Status);
END_FUNCTION

FUNCTION "FRK_CfgDef_DeclarationCell" : Void   // FC139, SCL
{ S7_Optimized_Access := 'TRUE' }
VERSION : 0.1
// stored: AutoNumber true, IsIECCheckEnabled false, SetENOAutomatically false, UDAEnableTagReadback false
   VAR_INPUT
      FieldIndex : Int;
   END_VAR
BEGIN

   "FRK_ConfigScratch".Entry := "FRK_ConfigScratch".Blank;
   CASE #FieldIndex OF
       1:
           "FRK_ConfigScratch".Entry.WriteKey := 'timeout';
           "FRK_ConfigScratch".Entry.WriteRevision := UDINT#1;
           "FRK_ConfigScratch".Entry.Item := WSTRING#'ParCfg/Timeout';
           "FRK_ConfigScratch".Entry.ConfigKind := 0;
           "FRK_ConfigScratch".Entry.ValueType := 3;
           "FRK_ConfigScratch".Entry.Writable := TRUE;
           "FRK_ConfigScratch".Entry.RequiresReady := TRUE;
           "FRK_ConfigScratch".Entry.HasMinimum := TRUE;
           "FRK_ConfigScratch".Entry.HasMaximum := TRUE;
           "FRK_ConfigScratch".Entry.Minimum := 1.0;
           "FRK_ConfigScratch".Entry.Maximum := 60000.0;
           "FRK_ConfigScratch".Entry.LabelKey := 'test.config.timeout';
           "FRK_ConfigScratch".Storage := 7;
           "FRK_ConfigScratch".Schema := 4;
           "FRK_ConfigScratch".Minimum := 1.0;
           "FRK_ConfigScratch".Maximum := 60000.0;
           "FRK_ConfigScratch".MaxLength := 0;
           "FRK_ConfigScratch".MinRead := 0;
           "FRK_ConfigScratch".MinWrite := 0;
       2:
           "FRK_ConfigScratch".Entry.WriteKey := 'preset';
           "FRK_ConfigScratch".Entry.WriteRevision := UDINT#2;
           "FRK_ConfigScratch".Entry.Item := WSTRING#'ParCfg/Preset';
           "FRK_ConfigScratch".Entry.ConfigKind := 0;
           "FRK_ConfigScratch".Entry.ValueType := 0;
           "FRK_ConfigScratch".Entry.Writable := TRUE;
           "FRK_ConfigScratch".Entry.RequiresReady := TRUE;
           "FRK_ConfigScratch".Entry.HasMinimum := TRUE;
           "FRK_ConfigScratch".Entry.HasMaximum := TRUE;
           "FRK_ConfigScratch".Entry.Minimum := 0.0;
           "FRK_ConfigScratch".Entry.Maximum := 1000.0;
           "FRK_ConfigScratch".Entry.LabelKey := 'test.config.preset';
           "FRK_ConfigScratch".Storage := 3;
           "FRK_ConfigScratch".Schema := 4;
           "FRK_ConfigScratch".Minimum := 0.0;
           "FRK_ConfigScratch".Maximum := 1000.0;
           "FRK_ConfigScratch".MaxLength := 0;
           "FRK_ConfigScratch".MinRead := 0;
           "FRK_ConfigScratch".MinWrite := 1;
       ELSE
           RETURN;
   END_CASE;
END_FUNCTION

FUNCTION "FRK_CfgDef_DeclarationCylinder" : Void   // FC131, SCL
{ S7_Optimized_Access := 'TRUE' }
VERSION : 0.1
// stored: AutoNumber true, IsIECCheckEnabled false, SetENOAutomatically false, UDAEnableTagReadback false
   VAR_INPUT
      FieldIndex : Int;
   END_VAR
BEGIN

   "FRK_ConfigScratch".Entry := "FRK_ConfigScratch".Blank;
   CASE #FieldIndex OF
       1:
           "FRK_ConfigScratch".Entry.WriteKey := 'timeout';
           "FRK_ConfigScratch".Entry.WriteRevision := UDINT#1;
           "FRK_ConfigScratch".Entry.Item := WSTRING#'ParCfg/Timeout';
           "FRK_ConfigScratch".Entry.ConfigKind := 0;
           "FRK_ConfigScratch".Entry.ValueType := 3;
           "FRK_ConfigScratch".Entry.Writable := TRUE;
           "FRK_ConfigScratch".Entry.RequiresReady := TRUE;
           "FRK_ConfigScratch".Entry.HasMinimum := TRUE;
           "FRK_ConfigScratch".Entry.HasMaximum := TRUE;
           "FRK_ConfigScratch".Entry.Minimum := 1.0;
           "FRK_ConfigScratch".Entry.Maximum := 60000.0;
           "FRK_ConfigScratch".Entry.LabelKey := 'test.config.timeout';
           "FRK_ConfigScratch".Storage := 7;
           "FRK_ConfigScratch".Schema := 4;
           "FRK_ConfigScratch".Minimum := 1.0;
           "FRK_ConfigScratch".Maximum := 60000.0;
           "FRK_ConfigScratch".MaxLength := 0;
           "FRK_ConfigScratch".MinRead := 0;
           "FRK_ConfigScratch".MinWrite := 0;
       2:
           "FRK_ConfigScratch".Entry.WriteKey := 'preset';
           "FRK_ConfigScratch".Entry.WriteRevision := UDINT#2;
           "FRK_ConfigScratch".Entry.Item := WSTRING#'ParCfg/Preset';
           "FRK_ConfigScratch".Entry.ConfigKind := 0;
           "FRK_ConfigScratch".Entry.ValueType := 0;
           "FRK_ConfigScratch".Entry.Writable := TRUE;
           "FRK_ConfigScratch".Entry.RequiresReady := TRUE;
           "FRK_ConfigScratch".Entry.HasMinimum := TRUE;
           "FRK_ConfigScratch".Entry.HasMaximum := TRUE;
           "FRK_ConfigScratch".Entry.Minimum := 0.0;
           "FRK_ConfigScratch".Entry.Maximum := 1000.0;
           "FRK_ConfigScratch".Entry.LabelKey := 'test.config.preset';
           "FRK_ConfigScratch".Storage := 3;
           "FRK_ConfigScratch".Schema := 4;
           "FRK_ConfigScratch".Minimum := 0.0;
           "FRK_ConfigScratch".Maximum := 1000.0;
           "FRK_ConfigScratch".MaxLength := 0;
           "FRK_ConfigScratch".MinRead := 0;
           "FRK_ConfigScratch".MinWrite := 1;
       ELSE
           RETURN;
   END_CASE;
END_FUNCTION

FUNCTION "FRK_CfgDef_DeclarationUnit" : Void   // FC164, SCL
{ S7_Optimized_Access := 'TRUE' }
VERSION : 0.1
// stored: AutoNumber true, IsIECCheckEnabled false, SetENOAutomatically false, UDAEnableTagReadback false
   VAR_INPUT
      FieldIndex : Int;
   END_VAR
BEGIN

